			etMunschExtruder :=  ET_MunschExtruder_eError;             (* Next step *)
		END_IF

	ET_MunschExtruder_eSetCMD:
		tonWatchdog(
			IN := TRUE,
			PT:= tTimeOutAir
		);

		IF tonWatchdog.Q
		THEN
			tonWatchdog(IN := FALSE);

			bExtruderAirOn := FALSE;

			udnErrorNo := 1;

			etMunschExtruder := ET_MunschExtruder_eError;             (* Next step *)

		ELSIF bExtruderAirOn
		THEN
			IF bExtruderAirOk
			THEN
				tonWatchdog(IN := FALSE);

				etMunschExtruder := ET_MunschExtruder_eSetMaterialTemp;              (* Next step *)
			END_IF
		ELSE
			Munsch.stMunschCmd.etCommand := ET_MUNSCH_CMD_STOPHEAT;

			tonWatchdog(IN := FALSE);

			etMunschExtruder := ET_MunschExtruder_eExecuteCMD;              (* Next step *)
		END_IF

	ET_MunschExtruder_eSetMaterialTemp:
		nWatchdog := nWatchdog + 1;

		Munsch.bLockedInterface := FALSE;

		fbMaterialTemp(
			bEnable := TRUE,
			bExecute := TRUE,
			nMaterialTemp := nMaterialTemp,
			nMinMaterialTemp := nMinMaterialTemp,
			nMaxMaterialTemp := nMaxMaterialTemp,
			Munsch := Munsch
		);

		IF (NOT fbMaterialTemp.bBusy
		     AND fbMaterialTemp.bError)
		     OR nWatchdog > 1000
		THEN
			fbMaterialTemp(
				bEnable := TRUE,
				bExecute := FALSE,
				Munsch := Munsch
			);

			udnErrorNo := 2;                     (* Error number *)

			etMunschExtruder := ET_MunschExtruder_eError;             (* Next step *)
		
		ELSIF NOT fbMaterialTemp.bBusy
			   AND  fbMaterialTemp.bDone
		THEN
			fbMaterialTemp(
				bEnable := TRUE,
				bExecute := FALSE,
				Munsch := Munsch
			);

			nWatchdog := 0;

			etMunschExtruder := ET_MunschExtruder_eSetAirTemp;             (* Next step *)

		END_IF;

		Munsch.bLockedInterface := TRUE;
		Munsch.bReadStatus := FALSE;

	ET_MunschExtruder_eSetAirTemp:
		nWatchdog := nWatchdog + 1;

		Munsch.bLockedInterface := FALSE;

		fbAirTemp(
			bEnable := TRUE,
			bExecute := TRUE,
			nAirTemp := nAirTemp,
			nMinAirTemp := nMinAirTemp,
			nMaxAirTemp := nMaxAirTemp,
			Munsch := Munsch
		);

		IF (NOT fbAirTemp.bBusy
		     AND fbAirTemp.bError)
		     OR nWatchdog > 1000
		THEN
			fbAirTemp(
				bEnable := TRUE,
				bExecute := FALSE,
				Munsch := Munsch
			);

			udnErrorNo := 3;                     (* Error number *)

			etMunschExtruder := ET_MunschExtruder_eError;             (* Next step *)

		ELSIF NOT fbAirTemp.bBusy
			   AND fbAirTemp.bDone
		THEN
			fbAirTemp(
				bEnable := TRUE,
				bExecute := FALSE,
				Munsch := Munsch
			);

			nWatchdog := 0;

			Munsch.stMunschCmd.etCommand := ET_MUNSCH_CMD_STARTHEAT;

			etMunschExtruder := ET_MunschExtruder_eExecuteCMD;             (* Next step *)
		
		END_IF;

		Munsch.bLockedInterface := TRUE;
		Munsch.bReadStatus := FALSE;

	ET_MunschExtruder_eExecuteCMD:
		nWatchdog := nWatchdog + 1;

		Munsch.bSendExe := TRUE;

		IF Munsch.bStringReceived
		THEN
			IF (bExtruderAirOn
			      AND Munsch.stMunschRes.etResponse = ET_MUNSCH_RES_STARTHEAT)
			     OR
			     (NOT bExtruderAirOn
			      AND Munsch.stMunschRes.etResponse = ET_MUNSCH_RES_STOPHEAT)
			THEN
				Munsch.bSendExe := FALSE;

				nWatchdog := 0;

				etMunschExtruder := ET_MunschExtruder_eSetREQ;              (* Next step *)

			END_IF

		ELSIF Munsch.bInterfaceError
			    OR nWatchdog > 1000
		THEN
			Munsch.bSendExe := FALSE;

			udnErrorNo := 4;                     (* Error number *)

			etMunschExtruder := ET_MunschExtruder_eError;              (* Next step *)

		END_IF

	ET_MunschExtruder_eSetREQ:
		Munsch.stMunschCmd.etCommand := ET_MUNSCH_CMD_REQHEATSTATUS;

		etMunschExtruder := ET_MunschExtruder_eExecuteREQ;              (* Next step *)

	ET_MunschExtruder_eExecuteREQ:
		nWatchdog := nWatchdog + 1;

		Munsch.bSendExe := TRUE;

		IF Munsch.bStringReceived
		THEN
			IF Munsch.stMunschRes.etResponse = ET_MUNSCH_RES_ACKHEATSTATUSON
			THEN
				Munsch.bHeat := TRUE;
				Munsch.bSendExe := FALSE;

				nWatchdog := 0;
				etMunschExtruder := ET_MunschExtruder_eDone;              (* Next step *)
			
			ELSIF Munsch.stMunschRes.etResponse = ET_MUNSCH_RES_ACKHEATSTATUSOFF
			THEN
				Munsch.bHeat := FALSE;
				Munsch.bSendExe := FALSE;

				nWatchdog := 0;
				etMunschExtruder := ET_MunschExtruder_eDone;              (* Next step *)

			END_IF

		ELSIF Munsch.bInterfaceError
			    OR nWatchdog > 1000
		THEN
			Munsch.bSendExe := FALSE;

			udnErrorNo := 5;                     (* Error number *)

			etMunschExtruder := ET_MunschExtruder_eError;              (* Next step *)

		END_IF

	ET_MunschExtruder_eError:
		bBusy := FALSE;						(* Command busy *)
		bError := TRUE;						(* Command error  *)

		etMunschExtruder := ET_MunschExtruder_eNoExecute;

	ET_MunschExtruder_eDone:
		bDone := TRUE;						(* Command done *)
		bBusy := FALSE;						(* Command busy *)

		etMunschExtruder := ET_MunschExtruder_eNoExecute;

	ET_MunschExtruder_eNoExecute:
		IF NOT bStart
		     AND NOT bStop
		THEN
			(* Reset outputs *)
			bDone := FALSE;						(* Command done *)
			bBusy := FALSE;						(* Command busy *)
			bError := FALSE;						(* Command error  *)

			nWatchdog := 0;
			Munsch.bLockedInterface := FALSE;

			Munsch.stMunschCmd.etCommand := ET_MUNSCH_CMD_NOCMD;
			Munsch.stMunschRes.etResponse := ET_MUNSCH_RES_NOCMD;

			etMunschExtruder := ET_MunschExtruder_eWaitExecute;
		END_IF
END_CASE;

END_FUNCTION_BLOCK

// ---- POUs/Tc3 Objects/ExternalHardware/Munsch/FB_MunschExtruder_MaterialTemp_1.TcPOU
FUNCTION_BLOCK FB_MunschExtruder_MaterialTemp_1
(*

The function block used to control set material temperature on munschs extruder

Constructor: 		Patryk Panylo
Company:		E. Riexinger GmbH
Date:			18.10.2015
Version:			1.00

Date:			Revision:		Who:				Comment
dd.mm.yyyy		x.xx			Initials			comment

*)
VAR_INPUT
	(* Input variables / Eingang Variablen *)
	bEnable						:BOOL;						(* Enable FB signal *)
	bExecute					:BOOL;						(* Execut the function block *)
	nMaterialTemp				:INT;						(* Material temperatur *)
	nMinMaterialTemp			:INT;						(* Minimal material temperatur *)
	nMaxMaterialTemp			:INT;						(* Maximal material temperatur *)
	nMaterialTempTolerance		:INT := 5;						(* Material temperatur tolerance*)
END_VAR
VAR_OUTPUT
	(* Output variables / Ausgang Variablen *)
	bMaterialTempAlarm			:BOOL;						(* Exceeded material temperature tolerance  *)
	bDone						:BOOL;						(* Program done *)
	bBusy						:BOOL;						(* Program busy *)
	bError						:BOOL;						(* Error *)
	udnErrorNo					:UDINT;
END_VAR
VAR_IN_OUT
	(* Input Output variables / Ausgang Variablen *)
	Munsch						:ST_MUNSCH_REF;
END_VAR
VAR
	(* Enummerations *)
	etMunschExtruder				:ET_MunschExtruder;

	(* Variables *)
	nWatchdog					:INT;

	(* References *)

	(* Interfaces *)

	(* Instances *)
	rtExecute						:R_TRIG;

END_VAR

IF NOT bEnable
THEN
	bDone := FALSE;					(* Program done *)
	bBusy := FALSE;                                  	(* Program not busy *)
	bError := FALSE;                                 	(* Program not error *)
	udnErrorNo := 0;                                 		(* Error number *)

	RETURN;
END_IF;

(* Wait for triger *)
rtExecute(CLK := bExecute);

(* Send command *)
CASE etMunschExtruder OF

	ET_MunschExtruder_eWaitExecute:
		IF rtExecute.Q
		THEN
			nWatchdog := 0;

			Munsch.bSetAirTemp := FALSE;
			Munsch.bSetMaterialTemp := TRUE;
			Munsch.bStartHeat := FALSE;
			Munsch.bStopHeat  := FALSE;
			Munsch.bStartExtruding := FALSE;
			Munsch.bStopExtruding  := FALSE;
			Munsch.bReadStatus := FALSE;

			etMunschExtruder := ET_MunschExtruder_eChkInterface;              (* Next step *)
		END_IF

	ET_MunschExtruder_eChkInterface:
		nWatchdog := nWatchdog + 1;

		IF NOT Munsch.bLockedInterface
		THEN
			bBusy := FALSE;                                     	(* Program not busy *)
			bError := FALSE;                         		(* Program not error *)
			udnErrorNo := 0;                         		(* Error number *)

			IF Munsch.bSetMaterialTemp
			THEN
				nWatchdog := 0;
				bDone:= FALSE;                               		(* Program done *)
				bBusy := TRUE;                                  	(* Program busy *)
	
				Munsch.bLockedInterface := TRUE;
				Munsch.bSendExe := FALSE;
	
				IF nMaterialTemp >= nMinMaterialTemp
				     AND nMaterialTemp <= nMaxMaterialTemp
				THEN
					etMunschExtruder := ET_MunschExtruder_eSetCMD;              (* Next step *)
				ELSE
					udnErrorNo := 1;
	
					etMunschExtruder := ET_MunschExtruder_eError;              (* Next step *)
				END_IF

			ELSE
				etMunschExtruder := ET_MunschExtruder_eError;             (* Next step *)
			END_IF

			Munsch.bSetMaterialTemp := FALSE;

		ELSIF nWatchdog > 1000
		THEN
			Munsch.bSetMaterialTemp := FALSE;

			etMunschExtruder := ET_MunschExtruder_eError;             (* Next step *)
		END_IF

	ET_MunschExtruder_eSetCMD:
		Munsch.stMunschCmd.etCommand := ET_MUNSCH_CMD_SETMATERIALTEMP;
		Munsch.stMunschCmd.nMaterialTemp := nMaterialTemp;

		etMunschExtruder := ET_MunschExtruder_eExecuteCMD;              (* Next step *)

	ET_MunschExtruder_eExecuteCMD:
		nWatchdog := nWatchdog + 1;

		Munsch.bSendExe := TRUE;

		IF Munsch.bStringReceived
		THEN
			IF Munsch.stMunschRes.etResponse = ET_MUNSCH_RES_SETMATERIALTEMP
			     AND Munsch.stMunschCmd.nMaterialTemp = Munsch.stMunschRes.nMaterialRefTemp
			THEN
				Munsch.bSendExe := FALSE;

				nWatchdog := 0;
				etMunschExtruder := ET_MunschExtruder_eSetREQ;              (* Next step *)
			END_IF

		ELSIF Munsch.bInterfaceError
			    OR nWatchdog > 1000
		THEN
			Munsch.bSendExe := FALSE;

			udnErrorNo := 2;                     (* Error number *)
			etMunschExtruder := ET_MunschExtruder_eError;              (* Next step *)
		END_IF

	ET_MunschExtruder_eSetREQ:
		Munsch.stMunschCmd.etCommand := ET_MUNSCH_CMD_REQMATERIALREFTEMP;

		etMunschExtruder := ET_MunschExtruder_eExecuteREQ;              (* Next step *)

	ET_MunschExtruder_eExecuteREQ:
		nWatchdog := nWatchdog + 1;

		Munsch.bSendExe := TRUE;

		IF Munsch.bStringReceived
		THEN
			IF Munsch.stMunschRes.etResponse = ET_MUNSCH_RES_REQMATERIALREFTEMP
			THEN
				Munsch.nMaterialRefTemp := Munsch.stMunschRes.nMaterialRefTemp;

				Munsch.bSendExe := FALSE;

				nWatchdog := 0;
				etMunschExtruder := ET_MunschExtruder_eDone;              (* Next step *)

			END_IF

		ELSIF Munsch.bInterfaceError
			    OR nWatchdog > 1000
		THEN
			Munsch.bSendExe := FALSE;

			udnErrorNo := 3;                     (* Error number *)
			etMunschExtruder := ET_MunschExtruder_eError;              (* Next step *)
		END_IF

	ET_MunschExtruder_eError:
		bBusy := FALSE;						(* Command busy *)
		bError := TRUE;						(* Command error  *)

		etMunschExtruder := ET_MunschExtruder_eNoExecute;

	ET_MunschExtruder_eDone:
		bDone := TRUE;						(* Command done *)
		bBusy := FALSE;						(* Command busy *)

		etMunschExtruder := ET_MunschExtruder_eNoExecute;

	ET_MunschExtruder_eNoExecute:
		IF NOT bExecute
		THEN
			(* Reset outputs *)
			bDone := FALSE;						(* Command done *)
			bBusy := FALSE;						(* Command busy *)
			bError := FALSE;						(* Command error  *)

			nWatchdog := 0;
			Munsch.bLockedInterface := FALSE;

			Munsch.stMunschCmd.etCommand := ET_MUNSCH_CMD_NOCMD;
			Munsch.stMunschRes.etResponse := ET_MUNSCH_RES_NOCMD;

			etMunschExtruder := ET_MunschExtruder_eWaitExecute;
		END_IF
END_CASE;

bMaterialTempAlarm := Munsch.nMaterialActTemp > Munsch.nMaterialRefTemp + nMaterialTempTolerance
					 OR Munsch.nMaterialActTemp > Munsch.nMaterialRefTemp - nMaterialTempTolerance;

END_FUNCTION_BLOCK

// ---- POUs/Tc3 Objects/ExternalHardware/Munsch/FB_MunschExtruder_ReadStatus_1.TcPOU
FUNCTION_BLOCK FB_MunschExtruder_ReadStatus_1
(*

The function block used to read status of Munsch extruder

Constructor: 		Patryk Panylo
Company:		E. Riexinger GmbH
Date:			13.10.2015
Version:			1.00

Date:			Revision:		Who:				Comment
dd.mm.yyyy		x.xx			Initials			comment

*)
VAR_INPUT
	(* Input variables / Eingang Variablen *)
	bEnable						:BOOL;						(* Enable FB signal *)
	bExecute					:BOOL;						(* Execute read status *)
	tReadStatus					:TIME := t#0ms;				(* Read current status *)
END_VAR
VAR_OUTPUT
	(* Output variables / Ausgang Variablen *)
	bDone						:BOOL;						(* Program done *)
	bBusy						:BOOL;						(* Program busy *)
	bError						:BOOL;						(* Error *)
	udnErrorNo					:UDINT;
END_VAR
VAR_IN_OUT
	(* Input Output variables / Ausgang Variablen *)
	Munsch						:ST_MUNSCH_REF;
END_VAR
VAR
	(* Enummerations *)
	etMunschExtruder				:ET_MunschExtruder;

	(* Variables *)
	bReadStatus					:BOOL;
	nReqCount					:INT;
	nWatchdog					:INT;

	(* References *)

	(* Interfaces *)

	(* Instances *)
	tonReadStatus				:TON;
	rtExecute						:R_TRIG;
	rtStart						:R_TRIG;
	rtStop						:R_TRIG;
END_VAR

IF NOT bEnable
THEN
	bDone := FALSE;					(* Program done *)
	bBusy := FALSE;                                  	(* Program not busy *)
	bError := FALSE;                                 	(* Program not error *)
	udnErrorNo := 0;                                 		(* Error number *)

	tonReadStatus(
		IN := FALSE,
	);

	RETURN;
END_IF;

rtStart(CLK := (tReadStatus > t#0ms
		       OR  (bExecute AND tReadStatus = t#0ms))
		       AND NOT Munsch.bLockedInterface);
rtStop(CLK := tReadStatus = t#0ms);

IF rtStop.Q
THEN
	Munsch.bReadStatus := FALSE;

ELSIF rtStart.Q
THEN
	Munsch.bReadStatus := TRUE;

	bDone := FALSE;					(* Program done *)
	bBusy := FALSE;                                  	(* Program not busy *)
	bError := FALSE;                                 	(* Program not error *)
	udnErrorNo := 0;                                 		(* Error number *)

	etMunschExtruder := ET_MunschExtruder_eWaitExecute;              (* Next step *)

END_IF

tonReadStatus(
	IN := Munsch.bReadStatus,
	PT := tReadStatus,
);

rtExecute(
	CLK := tonReadStatus.Q
);

(* Send command *)
CASE etMunschExtruder OF

	ET_MunschExtruder_eWaitExecute:
		bBusy := FALSE;                                     	(* Program not busy *)
		bError := FALSE;                         		(* Program not error *)
		udnErrorNo := 0;                         		(* Error number *)

		IF rtExecute.Q
		     AND NOT Munsch.bLockedInterface
		THEN
			nWatchdog := 0;
			bDone:= FALSE;                               		(* Program done *)
			bBusy := TRUE;                                  	(* Program busy *)

			nReqCount  := 0;
			Munsch.bLockedInterface := TRUE;
			Munsch.bSendExe := FALSE;

			etMunschExtruder := ET_MunschExtruder_eSetREQ;              (* Next step *)

		END_IF

	ET_MunschExtruder_eSetREQ:
		CASE nReqCount
		OF
			0: Munsch.stMunschCmd.etCommand := ET_MUNSCH_CMD_REQHEATSTATUS;
			    nReqCount := 1;
			1: Munsch.stMunschCmd.etCommand := ET_MUNSCH_CMD_REQEXTRUDERSTATUS;
			    nReqCount := 2;
			2: Munsch.stMunschCmd.etCommand := ET_MUNSCH_CMD_REQMATERIALREFTEMP;
			    nReqCount := 3;
			3: Munsch.stMunschCmd.etCommand := ET_MUNSCH_CMD_REQMATERIALACTTEMP;
			    nReqCount := 4;
			4: Munsch.stMunschCmd.etCommand := ET_MUNSCH_CMD_REQAIRREFTEMP;
			    nReqCount := 5;
			5: Munsch.stMunschCmd.etCommand := ET_MUNSCH_CMD_REQAIRACTTEMP;
			    nReqCount := 6;
			6: Munsch.stMunschCmd.etCommand := ET_MUNSCH_CMD_REQSTATUS;
				nReqCount := 0;
		END_CASE

		etMunschExtruder := ET_MunschExtruder_eExecuteREQ;              (* Next step *)

	ET_MunschExtruder_eExecuteREQ:
		nWatchdog := nWatchdog + 1;

		Munsch.bSendExe := TRUE;

		IF Munsch.bStringReceived
		THEN
			IF Munsch.stMunschRes.etResponse = ET_MUNSCH_RES_ACKHEATSTATUSON
			THEN
				Munsch.bHeat := TRUE;
				Munsch.bSendExe := FALSE;

				nWatchdog := 0;
				IF nReqCount > 0
				     AND Munsch.bReadStatus
				THEN
					etMunschExtruder := ET_MunschExtruder_eSetREQ;
				ELSE
					etMunschExtruder := ET_MunschExtruder_eDone;              (* Next step *)
				END_IF
			
			ELSIF Munsch.stMunschRes.etResponse = ET_MUNSCH_RES_ACKHEATSTATUSOFF
			THEN
				Munsch.bHeat := FALSE;
				Munsch.bSendExe := FALSE;

				nWatchdog := 0;
				IF nReqCount > 0
				    AND Munsch.bReadStatus
				THEN
					etMunschExtruder := ET_MunschExtruder_eSetREQ;
				ELSE
					etMunschExtruder := ET_MunschExtruder_eDone;              (* Next step *)
				END_IF

			ELSIF Munsch.stMunschRes.etResponse = ET_MUNSCH_RES_ACKEXTRUDERSTATUSON
			THEN
				Munsch.bExtruding := TRUE;
				Munsch.bSendExe := FALSE;

				nWatchdog := 0;
				IF nReqCount > 0
				    AND Munsch.bReadStatus
				THEN
					etMunschExtruder := ET_MunschExtruder_eSetREQ;
				ELSE
					etMunschExtruder := ET_MunschExtruder_eDone;              (* Next step *)
				END_IF
			
			ELSIF Munsch.stMunschRes.etResponse = ET_MUNSCH_RES_ACKEXTRUDERSTATUSOFF
			THEN
				Munsch.bExtruding := FALSE;
				Munsch.bSendExe := FALSE;

				nWatchdog := 0;
				IF nReqCount > 0
				     AND Munsch.bReadStatus
				THEN
					etMunschExtruder := ET_MunschExtruder_eSetREQ;
				ELSE
					etMunschExtruder := ET_MunschExtruder_eDone;              (* Next step *)
				END_IF

			ELSIF Munsch.stMunschRes.etResponse = ET_MUNSCH_RES_REQMATERIALREFTEMP
			THEN
				Munsch.nMaterialRefTemp := Munsch.stMunschRes.nMaterialRefTemp;
				Munsch.bSendExe := FALSE;

				nWatchdog := 0;
				IF nReqCount > 0
				     AND Munsch.bReadStatus
				THEN
					etMunschExtruder := ET_MunschExtruder_eSetREQ;
				ELSE
					etMunschExtruder := ET_MunschExtruder_eDone;              (* Next step *)
				END_IF

			ELSIF Munsch.stMunschRes.etResponse = ET_MUNSCH_RES_REQMATERIALACTTEMP
			THEN
				Munsch.nMaterialActTemp := Munsch.stMunschRes.nMaterialActTemp;
				Munsch.bSendExe := FALSE;

				nWatchdog := 0;
				IF nReqCount > 0
				     AND Munsch.bReadStatus
				THEN
					etMunschExtruder := ET_MunschExtruder_eSetREQ;
				ELSE
					etMunschExtruder := ET_MunschExtruder_eDone;              (* Next step *)
				END_IF

			ELSIF Munsch.stMunschRes.etResponse = ET_MUNSCH_RES_REQAIRREFTEMP
			THEN
				Munsch.nAirRefTemp := Munsch.stMunschRes.nAirRefTemp;
				Munsch.bSendExe := FALSE;

				nWatchdog := 0;
				IF nReqCount > 0
				     AND Munsch.bReadStatus
				THEN
					etMunschExtruder := ET_MunschExtruder_eSetREQ;
				ELSE
					etMunschExtruder := ET_MunschExtruder_eDone;              (* Next step *)
				END_IF

			ELSIF Munsch.stMunschRes.etResponse = ET_MUNSCH_RES_REQAIRACTTEMP
			THEN
				Munsch.nAirActTemp := Munsch.stMunschRes.nAirActTemp;
				Munsch.bSendExe := FALSE;

				nWatchdog := 0;
				IF nReqCount > 0
				     AND Munsch.bReadStatus
				THEN
					etMunschExtruder := ET_MunschExtruder_eSetREQ;
				ELSE
					etMunschExtruder := ET_MunschExtruder_eDone;              (* Next step *)
				END_IF

			ELSIF Munsch.stMunschRes.etResponse = ET_MUNSCH_RES_REQSTATUSHEATED
			THEN
				Munsch.bHeating := FALSE;
				Munsch.bHeated := TRUE;
				Munsch.bError := FALSE;
				Munsch.bSendExe := FALSE;

				nWatchdog := 0;
				IF nReqCount > 0
				     AND Munsch.bReadStatus
				THEN
					etMunschExtruder := ET_MunschExtruder_eSetREQ;
				ELSE
					etMunschExtruder := ET_MunschExtruder_eDone;              (* Next step *)
				END_IF

			ELSIF Munsch.stMunschRes.etResponse = ET_MUNSCH_RES_REQSTATUSHEATING
			THEN
				Munsch.bHeating := Munsch.bHeat;
				Munsch.bHeated := FALSE;
				Munsch.bError := FALSE;
				Munsch.bSendExe := FALSE;

				nWatchdog := 0;
				IF nReqCount > 0
				     AND Munsch.bReadStatus
				THEN
					etMunschExtruder := ET_MunschExtruder_eSetREQ;
				ELSE
					etMunschExtruder := ET_MunschExtruder_eDone;              (* Next step *)
				END_IF

			ELSIF Munsch.stMunschRes.etResponse = ET_MUNSCH_RES_REQSTATUSERROR
			THEN
				Munsch.bHeating := FALSE;
				Munsch.bHeated := FALSE;
				Munsch.bError := TRUE;
				Munsch.bSendExe := FALSE;

				nWatchdog := 0;
				IF nReqCount > 0
				     AND Munsch.bReadStatus
				THEN
					etMunschExtruder := ET_MunschExtruder_eSetREQ;
				ELSE
					etMunschExtruder := ET_MunschExtruder_eDone;              (* Next step *)
				END_IF

			END_IF

		ELSIF Munsch.bInterfaceError
 			    OR nWatchdog > 1000
		THEN
			Munsch.bSendExe := FALSE;

			udnErrorNo := 2;                     (* Error number *)

			etMunschExtruder := ET_MunschExtruder_eError;              (* Next step *)
		END_IF

	ET_MunschExtruder_eError:
		bBusy := FALSE;						(* Command busy *)
		bError := TRUE;						(* Command error  *)

		etMunschExtruder := ET_MunschExtruder_eNoExecute;

	ET_MunschExtruder_eDone:
		bDone := TRUE;						(* Command done *)
		bBusy := FALSE;						(* Command busy *)

		etMunschExtruder := ET_MunschExtruder_eNoExecute;

	ET_MunschExtruder_eNoExecute:
		IF tReadStatus > t#0ms
		THEN
			tonReadStatus(
				IN := FALSE,
				PT := tReadStatus,
			);
		END_IF

		IF NOT tonReadStatus.Q
		     OR (NOT bExecute AND tReadStatus = t#0ms)
		THEN
			(* Reset outputs *)
			bDone := FALSE;						(* Command done *)
			bBusy := FALSE;						(* Command busy *)
			bError := FALSE;						(* Command error  *)

			nWatchdog := 0;
			Munsch.bLockedInterface := FALSE;

			IF tReadStatus = t#0ms
			THEN
				Munsch.bReadStatus := FALSE;
			END_IF

			etMunschExtruder := ET_MunschExtruder_eWaitExecute;
		END_IF
END_CASE;

END_FUNCTION_BLOCK

// ---- POUs/Tc3 Objects/ExternalHardware/Munsch/FB_MUNSCH_EXTRUDER_REF_1.TcPOU
FUNCTION_BLOCK FB_MUNSCH_EXTRUDER_REF_1
VAR_INPUT
	bSendExe					:BOOL;						(* Send execute *)
	tSendPeriod					:TIME := t#0s;					(* Send data every period. If tSendPeriod is 0 then th function is not active *)
	bLockedInterface				:BOOL;						(* Locked interface *)
	bHeat						:BOOL;						(* Heat status ON = TRUE, OFF = FALSE *)
	bHeating						:BOOL;						(* Heating status ON = TRUE, OFF = FALSE *)
	bHeated						:BOOL;						(* Heated status ON = TRUE, OFF = FALSE *)
	bError						:BOOL;						(* Error ON = TRUE, OFF = FALSE *)
	bExtruding					:BOOL;						(* Extruder status ON = TRUE, OFF = FALSE *)
	nMaterialRefTemp			:INT;						(* Referenc material tamperature *)
	nMaterialActTemp				:INT;						(* Current material tamperature *)
	nAirRefTemp					:INT;						(* Referenc air tamperature *)
	nAirActTemp					:INT;						(* Current air tamperature *)
	stMunschCmd				:ST_MUNSCH_CMD_Data;
	stMunschRes					:ST_MUNSCH_RES_Data;
	bInterfaceReady				:BOOL;						(* Interface ready to use *)
	bInterfaceError				:BOOL;						(* Interface error *)
	bStringReceived				:BOOL;						(* String received *)
	bSetAirTemp					:BOOL;						(* Set air temperature *)
	bSetMaterialTemp			:BOOL;						(* Set material temperature *)
	bStartHeat					:BOOL;						(* Heat start *)
	bStopHeat					:BOOL;						(* Heat stop *)
	bStartExtruding				:BOOL;						(* Extruding start *)
	bStopExtruding				:BOOL;						(* Extruding start *)
	bReadStatus					:BOOL;						(* Enable read current status *)
	bExtrudingStop				:BOOL;						(* Extruding stop *)
	nExtrudingSpeed				:INT;						(* Extruding speed *)
END_VAR
VAR_OUTPUT

END_VAR
VAR_IN_OUT

END_VAR
VAR

END_VAR

;

END_FUNCTION_BLOCK

// ---- POUs/Tc3 Objects/ExternalHardware/Munsch/F_MunschCMD_1.TcPOU
FUNCTION F_MunschCMD_1 : STRING							(* Command to Munsch extruder *)
VAR_INPUT
	stMunschCmd			:ST_MUNSCH_CMD_Data;
END_VAR
VAR
	usnBaseMaterialTemp		:USINT := 160;					(* Base material temperature 160 °C *)
	usnBaseAirTemp			:USINT := 160;					(* Base air temperature 160 °C *)
END_VAR


CASE stMunschCmd.etCommand OF

	ET_MUNSCH_CMD_NOCMD:						F_MunschCMD := 'NoCmd';
	ET_MUNSCH_CMD_STARTHEAT:					F_MunschCMD := 'H1';
	ET_MUNSCH_CMD_STOPHEAT:					F_MunschCMD := 'H0';
	ET_MUNSCH_CMD_REQHEATSTATUS:			F_MunschCMD := 'h?';
	ET_MUNSCH_CMD_STARTEXTRUDER:			F_MunschCMD := 'R1';
	ET_MUNSCH_CMD_STOPEXTRUDER:				F_MunschCMD := 'R0';
	ET_MUNSCH_CMD_REQEXTRUDERSTATUS:		F_MunschCMD := 'r?';
	ET_MUNSCH_CMD_SETMATERIALTEMP:			F_MunschCMD := CONCAT('M', CHR(INT_TO_BYTE(MIN(MAX(stMunschCmd.nMaterialTemp - usnBaseMaterialTemp, 0), 240))));
	ET_MUNSCH_CMD_REQMATERIALREFTEMP:		F_MunschCMD := 'm?';
	ET_MUNSCH_CMD_REQMATERIALACTTEMP:		F_MunschCMD := 'n?';
	ET_MUNSCH_CMD_SETAIRTEMP:					F_MunschCMD := CONCAT('A', CHR(INT_TO_BYTE(MIN(MAX(stMunschCmd.nAirTemp - usnBaseAirTemp, 0), 240))));
	ET_MUNSCH_CMD_REQAIRREFTEMP:				F_MunschCMD := 'a?';
	ET_MUNSCH_CMD_REQAIRACTTEMP:				F_MunschCMD := 'b?';
	ET_MUNSCH_CMD_REQSTATUS:					F_MunschCMD := 's?';
ELSE
	F_MunschCMD := 'NoCmd';
END_CASE

END_FUNCTION

// ---- POUs/Tc3 Objects/ExternalHardware/Munsch/F_MunschRES_1.TcPOU
FUNCTION F_MunschRES_1 : ST_MUNSCH_RES_Data			(* Response from Munsch extruder *)
VAR_INPUT
	sResponse					:STRING	;
END_VAR
VAR
	usnBaseMaterialTemp		:USINT := 160;					(* Base material temperature 160 °C *)
	usnBaseAirTemp			:USINT := 160;					(* Base air temperature 160 °C *)
END_VAR


IF sResponse = 'H1'		THEN	F_MunschRES.etResponse := ET_MUNSCH_RES_STARTHEAT;
ELSIF sResponse = 'H0'	THEN	F_MunschRES.etResponse := ET_MUNSCH_RES_STOPHEAT;
ELSIF sResponse = 'h1'	THEN	F_MunschRES.etResponse := ET_MUNSCH_RES_ACKHEATSTATUSON;
ELSIF sResponse = 'h0'	THEN	F_MunschRES.etResponse := ET_MUNSCH_RES_ACKHEATSTATUSOFF;
ELSIF sResponse = 'R1'	THEN	F_MunschRES.etResponse := ET_MUNSCH_RES_STARTEXTRUDER;
ELSIF sResponse = 'R0'	THEN	F_MunschRES.etResponse := ET_MUNSCH_RES_STOPEXTRUDER;
ELSIF sResponse = 'r1'		THEN	F_MunschRES.etResponse := ET_MUNSCH_RES_ACKEXTRUDERSTATUSON;
ELSIF sResponse = 'r0'		THEN	F_MunschRES.etResponse := ET_MUNSCH_RES_ACKEXTRUDERSTATUSOFF;
ELSIF FIND(sResponse, 'M') = 1		THEN	F_MunschRES.etResponse := ET_MUNSCH_RES_SETMATERIALTEMP; F_MunschRES.nMaterialRefTemp := usnBaseMaterialTemp + ASC(DELETE(sResponse,LEN('M'), FIND(sResponse, 'M')));
ELSIF FIND(sResponse, 'm') = 1 		THEN	F_MunschRES.etResponse := ET_MUNSCH_RES_REQMATERIALREFTEMP; F_MunschRES.nMaterialRefTemp := usnBaseMaterialTemp + ASC(DELETE(sResponse,LEN('m'), FIND(sResponse, 'm')));
ELSIF FIND(sResponse, 'n') = 1 		THEN	F_MunschRES.etResponse := ET_MUNSCH_RES_REQMATERIALACTTEMP; F_MunschRES.nMaterialActTemp := usnBaseMaterialTemp + ASC(DELETE(sResponse,LEN('n'), FIND(sResponse, 'n')));
ELSIF FIND(sResponse, 'A') = 1		THEN	F_MunschRES.etResponse := ET_MUNSCH_RES_SETAIRTEMP; F_MunschRES.nAirRefTemp := usnBaseAirTemp + ASC(DELETE(sResponse,LEN('A'), FIND(sResponse, 'A')));
ELSIF FIND(sResponse, 'a') = 1		THEN	F_MunschRES.etResponse := ET_MUNSCH_RES_REQAIRREFTEMP; F_MunschRES.nAirRefTemp := usnBaseAirTemp + ASC(DELETE(sResponse,LEN('a'), FIND(sResponse, 'a')));
ELSIF FIND(sResponse, 'b') = 1		THEN	F_MunschRES.etResponse := ET_MUNSCH_RES_REQAIRACTTEMP; F_MunschRES.nAirActTemp := usnBaseAirTemp + ASC(DELETE(sResponse,LEN('b'), FIND(sResponse, 'b')));
ELSIF sResponse = 's1'	THEN	F_MunschRES.etResponse := ET_MUNSCH_RES_REQSTATUSHEATED;
ELSIF sResponse = 's0'	THEN	F_MunschRES.etResponse := ET_MUNSCH_RES_REQSTATUSHEATING;
ELSIF sResponse = 'sE'	THEN	F_MunschRES.etResponse := ET_MUNSCH_RES_REQSTATUSERROR;
ELSIF sResponse = 'ER' 	THEN	F_MunschRES.etResponse := ET_MUNSCH_RES_CMDERROR;
ELSE F_MunschRES.etResponse := ET_MUNSCH_RES_NOCMD;
END_IF

END_FUNCTION

// ---- POUs/Tc3 Objects/ExternalHardware/Periphery/FB_PERIPHERY_REF_1.TcPOU
FUNCTION_BLOCK FB_PERIPHERY_REF_1
VAR_INPUT

END_VAR
VAR_OUTPUT

END_VAR
VAR_IN_OUT

END_VAR
VAR

END_VAR

;

END_FUNCTION_BLOCK

// ---- POUs/Tc3 Objects/ExternalHardware/YASKAWA/FB_YASKAWA_Controller_1.TcPOU
FUNCTION_BLOCK FB_YASKAWA_Controller_1
(*

The function block used to control axis.

Constructor: 		Patryk Panylo
Company:		E. Riexinger GmbH
Date:			20.06.2018
Version:			1.00

Date:			Revision:		Who:				Comment
dd.mm.yyyy		x.xx			Initials			comment

*)
VAR_INPUT
	(* Input variables / Eingang Variablen *)
	bEnable						:BOOL;						(* Signal FB enable *)
	etMachineMode				:ET_MachineMode;			(* Machine mode *)
	etMachineState				:ET_MachineState;			(* Machine state *)
	bDrivesOn					:BOOL;						(* Enable the drives *)
	bMoveOn					:BOOL;						(* Enable the move enable *)
	bReset						:BOOL;						(* Signal reset *)
	bExeReset					:BOOL;						(* Execute auto reset *)
	lrOverride					:LREAL;						(* Override 100% percent *)
END_VAR
VAR_OUTPUT
	(* Output variables / Ausgang Variablen *)
	bStatus						:BOOL;						(* Feedback *)
	bStatusDelay					:BOOL;						(* Feedback delay *)
	bReseted					:BOOL;						(* Reset completed *)
	bError						:BOOL;						(* Controller error *)
	udnErrorNo					:UDINT;						(* Error number *)
	bInHome						:BOOL;						(* In home *)
	bNotMoving					:BOOL;						(* Status of moving *)
	bNotInCrashAreaMachine		:BOOL;						(* Status not in crash area *)
END_VAR
VAR_IN_OUT
	(* Input Output variables / Ausgang Variablen *)
	Yaskawa					:ST_YASKAWA_REF;				(* The YASKAWA_REF data type  is an interface between the PLC and the YASKAWA and contains axis information *)
END_VAR
VAR
	(* Enummerations *)

	(* Variables *)
	tStatusDelay					:TIME := t#1s;					(* Status delay time *)

	bFirstTime					:BOOL;

	(* References *)

	(* Interfaces *)

	(* Instances *)
	fbPower						:FB_YASKAWA_Power;		(* The function block is used to enable for an axis *)
	tonStatusDelay				:TON;						(* Delay controller enabled status *)
	fbReset						:FB_YASKAWA_Reset;			(* An axis reset is carried out with the function block *)

END_VAR


IF NOT bEnable							(* Signal FB enable *)
THEN
	bStatus := FALSE;						(* Feedback *)
	bStatusDelay := FALSE;				(* Feedback *)
	bError := FALSE;						(* Controller error *)
	udnErrorNo := 0;						(* Error number *)

	bFirstTime := FALSE;
	RETURN;
END_IF

IF NOT bFirstTime
THEN

	bFirstTime := TRUE;
END_IF;

A_Power();
A_Reset();
A_Error();

(* In home *)
bInHome := Yaskawa.stYaskawaToPlc.bInHome;

(* Status not moving *)
bNotMoving := Yaskawa.stYaskawaToPlc.bNotMoving;

(* Status not in crash area *)
bNotInCrashAreaMachine := Yaskawa.stYaskawaToPlc.bNotInCrashAreaMachine;

ACTION A_Error:

bError := fbReset.bError
	         OR fbPower.bError;
END_ACTION

ACTION A_Power:

fbPower(
	bEnable := TRUE,
	bAutoHand := etMachineMode = ET_MachineMode_eHome
			         OR etMachineMode = ET_MachineMode_eStepping
			         OR etMachineMode = ET_MachineMode_eAutomatic
					 OR etMachineMode = ET_MachineMode_eMaintenance,
	bDrivesOn :=  bDrivesOn,
	bMoveOn := bMoveOn,
	lrOverride := lrOverride,
	Yaskawa := Yaskawa
 );

tonStatusDelay(
	IN := fbPower.bStatus,
	PT := SEL(etMachineMode = ET_MachineMode_eManual, tStatusDelay, t#0ms),
	Q => bStatusDelay
);
END_ACTION

ACTION A_Reset:

fbReset(
	bExecute := bReset
	            	     XOR bExeReset,
	Yaskawa := Yaskawa,
	bDone => bReseted
);
END_ACTION

END_FUNCTION_BLOCK

// ---- POUs/Tc3 Objects/ExternalHardware/YASKAWA/FB_YASKAWA_Power_1.TcPOU
FUNCTION_BLOCK FB_YASKAWA_Power_1
(*

The function block used to enable drives for an yaskawa

Constructor: 		Patryk Panylo
Company:		E. Riexinger GmbH
Date:			20.06.2018
Version:			1.00

Date:			Revision:		Who:				Comment

*)
VAR_INPUT
	(* Input variables / Eingang Variablen *)
	bEnable						:BOOL;			(* Signal FB enable *)
	bAutoHand					:BOOL;			(* Auto := TRUE, Hand := FALSE *)
	bDrivesOn					:BOOL;			(* Enable the drives *)
	bMoveOn					:BOOL;			(* Enable the move enable *)
	lrOverride					:LREAL;			(* Velocity override in % for all motion commands. (0 <= Override <= 100.0) *)
END_VAR
VAR_OUTPUT
	(* Output variables / Ausgang Variablen *)
	bStatus						:BOOL;			(* Status = TRUE indicates that the axis is ready for operation. *)
	bError						:BOOL;			(* Error *)
	udnErrorNo					:UDINT;			(* Error number *)
	sErrorMsg					:STRING; 		(* Error message *)
END_VAR
VAR_IN_OUT
	(* Input Output variables / Ausgang Variablen *)
	Yaskawa					:ST_YASKAWA_REF;				(* The YASKAWA_REF data type  is an interface between the PLC and the YASKAWA and contains axis information *)
END_VAR
VAR
	(* Enummerations *)

	(* Variables *)
	tStatusDelay 					:TIME := t#300ms;

	(* References *)

	(* Interfaces *)

	(* Instances *)
	tonStatusDelay				:TON;
END_VAR


IF NOT bEnable
THEN
	Yaskawa.stPlcToYaskawa.bExternalServoOn := FALSE;                   		 (* Switch on *)
	tonStatusDelay(IN := FALSE,
				    PT := tStatusDelay);
ELSE

	IF NOT bDrivesOn
	     OR Yaskawa.stYaskawaToPlc.bAlarmErrorOccured
	THEN
		Yaskawa.stPlcToYaskawa.bCallMasterJob := FALSE;
		Yaskawa.stPlcToYaskawa.bExternalStart := FALSE;
		Yaskawa.stPlcToYaskawa.bExternalHold := FALSE;
		Yaskawa.stPlcToYaskawa.bExternalServoOn := FALSE;						 (* Switch on *)
		Yaskawa.stPlcToYaskawa.bExternalServoOffEStop := TRUE;                   		 (* Switch off *)
		Yaskawa.stPlcToYaskawa.bExternalServoOffHoldStop := FALSE;                   		 (* Switch off *)
	ELSE
		IF bAutoHand			(* Auto *)
		THEN
			IF bMoveOn
			     AND Yaskawa.stYaskawaToPlc.bRemoteModeSelected
			THEN
				Yaskawa.stPlcToYaskawa.bExternalServoOn := TRUE;                   				 (* Switch on *)
				Yaskawa.stPlcToYaskawa.bExternalServoOffEStop := FALSE;                   		 (* Switch off *)
				Yaskawa.stPlcToYaskawa.bExternalServoOffHoldStop := FALSE;                   		 (* Switch off *)
			ELSE
				Yaskawa.stPlcToYaskawa.bExternalServoOn := FALSE;                   				(* Switch on *)
				Yaskawa.stPlcToYaskawa.bExternalServoOffEStop := FALSE;                   		(* Switch off *)
				Yaskawa.stPlcToYaskawa.bExternalServoOffHoldStop := TRUE;				(* Switch off *)
			END_IF
		ELSE				(* Manual *)
			Yaskawa.stPlcToYaskawa.bCallMasterJob := FALSE;
			Yaskawa.stPlcToYaskawa.bExternalStart := FALSE;
			Yaskawa.stPlcToYaskawa.bExternalHold := FALSE;
			Yaskawa.stPlcToYaskawa.bExternalServoOn := FALSE;						(* Switch on *)
			Yaskawa.stPlcToYaskawa.bExternalServoOffEStop := FALSE;                   		(* Switch off *)
			Yaskawa.stPlcToYaskawa.bExternalServoOffHoldStop := FALSE;				(* Switch off *)
		END_IF
	END_IF;
END_IF;

Yaskawa.stPlcToYaskawa.nOverride := LREAL_TO_INT(LIMIT(0,lrOverride,100));

tonStatusDelay(IN := Yaskawa.stYaskawaToPlc.bServoIsOn,		(* Control enabled *)
			   PT := tStatusDelay);
bStatus := tonStatusDelay.Q;

END_FUNCTION_BLOCK

// ---- POUs/Tc3 Objects/ExternalHardware/YASKAWA/FB_YASKAWA_REF_1.TcPOU
FUNCTION_BLOCK FB_YASKAWA_REF_1
VAR_INPUT
	stYaskawaToPlc				:ST_YASKAWATOPLC;
	stPlcToYaskawa				:ST_PLCTOYASKAWA;

	stRobotToPlc					AT %I*:ST_ROBOTTOPLC;
	stPlcToRobot					AT %Q*:ST_PLCTOROBOT;
END_VAR
VAR_OUTPUT

END_VAR
VAR_IN_OUT

END_VAR
VAR

END_VAR

;

END_FUNCTION_BLOCK

// ---- POUs/Tc3 Objects/ExternalHardware/YASKAWA/FB_YASKAWA_Reset_1.TcPOU
FUNCTION_BLOCK FB_YASKAWA_Reset_1
(*

The function block used to reset the yaskawa message.

Constructor: 		Patryk Panylo
Company:		E. Riexinger GmbH
Date:			20.06.2018
Version:			1.00

Date:			Revision:		Who:				Comment

*)
VAR_INPUT
	(* Input variables / Eingang Variablen *)
	bExecute					:BOOL;		(* Execut the function block *)
	bExtReset					:BOOL;
END_VAR
VAR_OUTPUT
	(* Output variables / Ausgang Variablen *)
	bDone						:BOOL;			(* Program done. *)
	bBusy						:BOOL;			(* Program busy *)
	bError						:BOOL;			(* Error *)
	udnErrorNo					:UDINT;			(* Error number *)
	sErrorMsg					:STRING; 		(* Error message *)
END_VAR
VAR_IN_OUT
	(* Input Output variables / Ausgang Variablen *)
	Yaskawa					:ST_YASKAWA_REF;				(* The YASKAWA_REF data type  is an interface between the PLC and the YASKAWA and contains axis information *)
END_VAR
VAR
	(* Enummerations *)

	(* Variables *)

	(* References *)

	(* Interfaces *)

	(* Instances *)
	rtExecute						:R_TRIG;
	rtExtReset					:R_TRIG;
	rtDrivesOn					:R_TRIG;

END_VAR


rtExecute(CLK := bExecute
			      AND Yaskawa.stYaskawaToPlc.bAlarmErrorOccured);
rtDrivesOn(CLK := Yaskawa.stYaskawaToPlc.bServoIsOn
	   		        AND Yaskawa.stPlcToYaskawa.bExternalServoOn);

IF rtExecute.Q
     OR (rtDrivesOn.Q
	    AND Yaskawa.stYaskawaToPlc.bAlarmErrorOccured)
THEN
	bBusy := TRUE;
	Yaskawa.stPlcToYaskawa.bAlarmReset := TRUE;

ELSIF Yaskawa.stPlcToYaskawa.bAlarmReset
	   AND NOT Yaskawa.stYaskawaToPlc.bAlarmErrorOccured
THEN
	bBusy := FALSE;
	Yaskawa.stPlcToYaskawa.bAlarmReset := FALSE;
END_IF;

bDone := bExecute
		AND NOT bBusy
		AND NOT Yaskawa.stYaskawaToPlc.bAlarmErrorOccured;        (* Error *)

END_FUNCTION_BLOCK

// ---- POUs/Tc3 Objects/ExternalHardware/YASKAWA/FB_YASKAWA_StartPrg_1.TcPOU
FUNCTION_BLOCK FB_YASKAWA_StartPrg_1
(*

The function block used to start kuka

Constructor: 		Patryk Panylo
Company:		E. Riexinger GmbH
Date:			18.11.2016
Version:			1.00

Date:			Revision:		Who:				Comment

*)
VAR_INPUT
	(* Input variables / Eingang Variablen *)
	bEnable						:BOOL;			(* Signal FB enable *)
	bReset						:BOOL;			(* Signal reset *)
	bAutoHand					:BOOL;			(* Auto := TRUE, Hand := FALSE *)
	bStart						:BOOL;			(* Start program *)
	bStop						:BOOL;			(* Stop program *)
	nPrgNo						:INT;			(* Program number *)
END_VAR
VAR_OUTPUT
	(* Output variables / Ausgang Variablen *)
	bRunning					:BOOL;						(* Program running *)
	bDone						:BOOL;						(* Program done *)
	bBusy						:BOOL;						(* Program busy *)
	bError						:BOOL;						(* Error *)
	udnErrorNo					:UDINT;
END_VAR
VAR_IN_OUT
	(* Input Output variables / Ausgang Variablen *)
	Yaskawa					:ST_YASKAWA_REF;				(* The YASKAWA_REF data type  is an interface between the PLC and the YASKAWA and contains axis information *)
END_VAR
VAR
	(* Enummerations *)
	etYaskawaStart				:ET_YaskawaStart;

	(* Variables *)
	bFirstTime					:BOOL;

	nWatchdog					:INT;

	(* References *)

	(* Interfaces *)

	(* Instances *)
	rtStart						:R_TRIG;
	rtStop						:R_TRIG;
	rtReset						:R_TRIG;
	tonWatchdog					:TON;

END_VAR


IF NOT bEnable
THEN
	bDone := FALSE;					(* Program done *)
	bBusy := FALSE;                                  	(* Program not busy *)
	bError := FALSE;                                 	(* Program not error *)
	udnErrorNo := 0;                                 		(* Error number *)

	Yaskawa.stPlcToYaskawa.bCallMasterJob := FALSE;
	Yaskawa.stPlcToYaskawa.bExternalStart := FALSE;
	Yaskawa.stPlcToYaskawa.bExternalHold := FALSE;

	RETURN;
END_IF;

IF NOT bFirstTime
THEN
	tonWatchdog(IN := FALSE);

	Yaskawa.stPlcToYaskawa.bCallMasterJob := FALSE;
	Yaskawa.stPlcToYaskawa.bExternalStart := FALSE;
	Yaskawa.stPlcToYaskawa.bExternalHold := FALSE;

	etYaskawaStart := ET_YaskawaStart_eWaitExecute;              (* Next step *)

	bFirstTime := TRUE;
END_IF

rtReset(CLK := bReset);

IF rtReset.Q
     AND bError
THEN
	bError := FALSE;

	tonWatchdog(IN := FALSE);

	Yaskawa.stPlcToYaskawa.bCallMasterJob := FALSE;
	Yaskawa.stPlcToYaskawa.bExternalStart := FALSE;
	Yaskawa.stPlcToYaskawa.bExternalHold := FALSE;

	etYaskawaStart := ET_YaskawaStart_eWaitExecute;              (* Next step *)
END_IF

(* Wait for triger *)
rtStart(
	CLK := bStart
);

IF rtStart.Q
     AND Yaskawa.stYaskawaToPlc.bServoIsOn
     AND NOT Yaskawa.stYaskawaToPlc.bAlarmErrorOccured
THEN
	Yaskawa.stPlcToYaskawa.bCallMasterJob := FALSE;
	Yaskawa.stPlcToYaskawa.bExternalStart := FALSE;
	Yaskawa.stPlcToYaskawa.bExternalHold := FALSE;

	etYaskawaStart := ET_YaskawaStart_eWaitExecute;              (* Next step *)

END_IF

rtStop(
	CLK := bStop
);

IF rtStop.Q
     OR Yaskawa.stYaskawaToPlc.bAlarmErrorOccured
THEN
	Yaskawa.stPlcToYaskawa.bCallMasterJob := FALSE;
	Yaskawa.stPlcToYaskawa.bExternalStart := FALSE;
	Yaskawa.stPlcToYaskawa.bExternalHold := Yaskawa.stYaskawaToPlc.bOperatingRunning
										     AND NOT Yaskawa.stYaskawaToPlc.bAlarmErrorOccured;

	etYaskawaStart := ET_YaskawaStart_eWaitExecute;              (* Next step *)

END_IF

bRunning := Yaskawa.stYaskawaToPlc.bOperatingRunning;
Yaskawa.stPlcToYaskawa.nPrgNo := nPrgNo;

(* Send command *)
CASE etYaskawaStart OF

	ET_YaskawaStart_eWaitExecute:
		bBusy := FALSE;                                     	(* Program not busy *)
		bError := FALSE;                         		(* Program not error *)
		udnErrorNo := 0;                         		(* Error number *)

		IF rtStart.Q
     		     AND bAutoHand			(* Automatic *)
		     AND NOT bStop
		THEN
			nWatchdog := 0;
			bDone:= FALSE;                               		(* Program done *)
			bBusy := TRUE;                                  	(* Program busy *)

			tonWatchdog(IN := FALSE);

			Yaskawa.stPlcToYaskawa.bCallMasterJob := FALSE;
			Yaskawa.stPlcToYaskawa.bExternalStart := FALSE;
			Yaskawa.stPlcToYaskawa.bExternalHold := FALSE;

			IF Yaskawa.stYaskawaToPlc.bHold
			THEN
				etYaskawaStart := ET_YaskawaStart_eExternalStart;              (* Next step *)
			ELSE
				etYaskawaStart := ET_YaskawaStart_eCallMasterJob;              (* Next step *)
			END_IF
		END_IF

	ET_YaskawaStart_eCallMasterJob:
		nWatchdog := nWatchdog + 1;

		Yaskawa.stPlcToYaskawa.bCallMasterJob := TRUE;

		IF Yaskawa.stYaskawaToPlc.bTopMasterJob
		     AND Yaskawa.stYaskawaToPlc.bServoIsOn
		     AND NOT Yaskawa.stYaskawaToPlc.bAlarmErrorOccured
		THEN
			nWatchdog := 0;

			Yaskawa.stPlcToYaskawa.bCallMasterJob := FALSE;

			etYaskawaStart := ET_YaskawaStart_eExternalStart;              (* Next step *)

		ELSIF Yaskawa.stYaskawaToPlc.bAlarmErrorOccured
			    OR nWatchdog > 1000
		THEN
			Yaskawa.stPlcToYaskawa.bCallMasterJob := FALSE;
			
			udnErrorNo := 1;                     (* Error number *)
			
			etYaskawaStart := ET_YaskawaStart_eError;              (* Next step *)

		END_IF

	ET_YaskawaStart_eExternalStart:
		nWatchdog := nWatchdog + 1;

		Yaskawa.stPlcToYaskawa.bExternalStart := TRUE;

		IF Yaskawa.stYaskawaToPlc.bOperatingRunning
		     AND Yaskawa.stYaskawaToPlc.bServoIsOn
		     AND NOT Yaskawa.stYaskawaToPlc.bPrgDone
		     AND NOT Yaskawa.stYaskawaToPlc.bAlarmErrorOccured
		THEN
			nWatchdog := 0;

			Yaskawa.stPlcToYaskawa.bExternalStart := FALSE;

			etYaskawaStart := ET_YaskawaStart_eWfPrgDone;              (* Next step *)

		ELSIF Yaskawa.stYaskawaToPlc.bAlarmErrorOccured
			    OR nWatchdog > 1000
		THEN
			Yaskawa.stPlcToYaskawa.bExternalStart := FALSE;
			
			udnErrorNo := 2;                     (* Error number *)

			etYaskawaStart := ET_YaskawaStart_eError;              (* Next step *)

		END_IF

	ET_YaskawaStart_eWfPrgDone:
		IF (Yaskawa.stYaskawaToPlc.bInHome
		     OR Yaskawa.stYaskawaToPlc.bNotInCrashAreaMachine)
		    AND Yaskawa.stYaskawaToPlc.bPrgDone
	     	    AND NOT Yaskawa.stYaskawaToPlc.bAlarmErrorOccured
		THEN
			Yaskawa.stPlcToYaskawa.bCallMasterJob := FALSE;;
			Yaskawa.stPlcToYaskawa.bExternalStart := FALSE;

			etYaskawaStart := ET_YaskawaStart_eDone;              (* Next step *)

		ELSIF Yaskawa.stYaskawaToPlc.bAlarmErrorOccured
		THEN
			Yaskawa.stPlcToYaskawa.bCallMasterJob := FALSE;;
			Yaskawa.stPlcToYaskawa.bExternalStart := FALSE;

			udnErrorNo := 3;                     (* Error number *)

			etYaskawaStart := ET_YaskawaStart_eError;              (* Next step *)

		END_IF

	ET_YaskawaStart_eError:
		bBusy := FALSE;						(* Command busy *)
		bError := TRUE;						(* Command error  *)

		etYaskawaStart := ET_YaskawaStart_eNoExecute;

	ET_YaskawaStart_eDone:
		bDone := TRUE;						(* Command done *)
		bBusy := FALSE;						(* Command busy *)

		etYaskawaStart := ET_YaskawaStart_eNoExecute;

	ET_YaskawaStart_eNoExecute:
		IF NOT bStart
		THEN
			(* Reset outputs *)
			bDone := FALSE;						(* Command done *)
			bBusy := FALSE;						(* Command busy *)
			bError := FALSE;						(* Command error  *)

			nWatchdog := 0;

			etYaskawaStart := ET_YaskawaStart_eWaitExecute;
		END_IF
END_CASE;

END_FUNCTION_BLOCK

// ---- POUs/Tc3 Objects/File/CSV/FB_FileCSVHandler.TcPOU
FUNCTION_BLOCK FB_FileCSVHandler
(*

This function block is used to read and write datas into/from csv file.
None of the field value is containing any non-printing control characters like line feed, carriage return, quotation marks, semicolon... 

Constructor: 		Patryk Panylo
Company:			E. Riexinger GmbH
Date:				05.04.2019
Version:			1.00

Date:			Revision:		Who:				Comment
dd.mm.yyyy		x.xx			Initials			comment

*)

VAR_INPUT
	bEnable						:BOOL := FALSE;				(* Enable FB *)
	sNetID						:T_AmsNetID	:= '';			(* TwinCAT Net ID *)
	bExecute					:BOOL := FALSE;				(* Execute operation *)
	sFilePath					:T_MaxString := '';			(* File path *)
	sFileName					:T_MaxString := '';			(* File name *)
	bCommaSeparator				:BOOL := FALSE;				(* Enable comma csv separator *)
	dwOpenMode					:DWORD;				(*
															FOPEN_MODEREAD (16#0001)	"r": Opens for reading. If the file does not exist or cannot be found, the call fails.
															FOPEN_MODEWRITE (16#0002) "w": Opens an empty file for writing. If the given file exists, its contents are destroyed.
															FOPEN_MODEAPPEND (16#0004) "a": Opens for writing at the end of the file (appending) without removing the EOF marker before writing new data to the file; creates the file first if it doesn’t exist.
															FOPEN_MODEREAD OR FOPEN_MODEPLUS (16#0008) "r+": Opens for reading and writing. The file must exist.
															FOPEN_MODEWRITE OR FOPEN_MODEPLUS (16#0008) "w+": Opens an empty file for both reading and writing. If the given file exists, its contents are destroyed.
															FOPEN_MODEAPPEND OR FOPEN_MODEPLUS (16#0008)	 "a+": Opens for reading and appending; the appending operation includes the removal of the EOF marker before new data is written to the file and the EOF marker is restored after writing is complete; creates the file first if it doesn’t exist.
															When a file is opened with the "a" or "a+" access type, all write operations occur at the end of the file. The file pointer can be repositioned using FB_FileSeek, but is always moved back to the end of the file before any write operation is carried out. Thus, existing data cannot be overwritten.
															
															FOPEN_MODEBINARY (16#0010) "b": Open in binary (untranslated) mode.
															FOPEN_MODETEXT (16#0020) "t": Open in text (translated) mode.
														*)
	arsWriteRecords				:ARRAY[0..GVL_CSV.MAX_CSV_ROWS, 0..GVL_CSV.MAX_CSV_COLUMNS ] OF STRING(GVL_CSV.MAX_CSV_FIELD_LENGTH);			(* Write records *)
	udnRowUsingMax				:UDINT;						(* Maximal number of using rows *)
	udnColumnUsingMax			:UDINT;						(* Maximal number of using columns *)																				
	tTimeout					:TIME := T#1S;				(* States the time before the function is cancelled *)
END_VAR
VAR_OUTPUT
	arsReadRecords				:ARRAY[0..GVL_CSV.MAX_CSV_ROWS, 0..GVL_CSV.MAX_CSV_COLUMNS ] OF STRING(GVL_CSV.MAX_CSV_FIELD_LENGTH);			(* Read records *)																										
	bBusy						:BOOL;					(* Program busy *)
	bDone						:BOOL;					(* Program done *)
	bError						:BOOL;					(* Program error *)
	udnErrNo					:UDINT;					(* Error number *)
END_VAR
VAR_IN_OUT

END_VAR
VAR
	(* Enummerations *)
	etCSVState					:ET_CSV_State := ET_CSV_State_eWaitExecute;
	
	(* Variables *)
	bFirstTime					:BOOL;					(* First PLC cycle *)

	dwModeCache					:DWORD;					(* Contains the mode in which the file is to be opened *)
	sPathName					:STRING;				(* Contains the path and filename for the file to be opened *)
	hFileHandle					:UINT;					(* File handle *)

	udnWriteCounter				:UDINT;
	udnReadCounter				:UDINT;

	udnRowCounter				:UDINT;
	udnColumnCounter			:UDINT;
	
	sCSVLine					:T_MaxString := '';		(* Single CSV text line (row, record), we are using string as record buffer (your are able to see created fields) *)
	sCSVField					:T_MaxString := '';		(* Single CSV field value (column, record field) *)
	
	(* Instances *)
	fbCreateDir					:FB_CreateDir;			(* Create direction *)
	
	fbFileOpen					:FB_FileOpen;			(* File open *)
	fbFileClose					:FB_FileClose;			(* File close *)

	fbFilePuts					:FB_FilePuts;			(* Writes one record (line) *)
	fbWriter					:FB_CSVMemBufferWriter;	(* Helper function block used to create CSV data bytes (single record line) *)
	
	fbFileGets					:FB_FileGets;			(* Reads one record (line) *)
	fbReader					:FB_CSVMemBufferReader;	(* Helper function block used to parse CSV data bytes (single record line) *)
END_VAR
VAR CONSTANT
	sFileSuffix					:STRING(5) := 'csv';
END_VAR

IF NOT bEnable				(* Enable FB *)
THEN
	bFirstTime := FALSE;		(* First PLC cycle *)
	bBusy := FALSE;			(* Program busy *)
	bDone := FALSE;			(* Program done *)
	bError := FALSE;			(* Program error *)
	udnErrNo := 0;				(* Error number *)
	RETURN;
END_IF

IF NOT bFirstTime
THEN
	IF bCommaSeparator
	THEN
		DEFAULT_CSV_FIELD_SEP := 16#2C;			(* Comma ASCII code *)
	ELSE
		DEFAULT_CSV_FIELD_SEP := 16#3B;			(* Semicolon ASCII code *)
	END_IF

	etCSVState := ET_CSV_State_eWaitExecute;

	bFirstTime := TRUE;
END_IF


(* Sequence state for open, read/write and close the file *)
CASE etCSVState
OF
	ET_CSV_State_eWaitExecute:
		IF bExecute
		THEN				
			fbCreateDir(
				sNetId:= sNetID,
				sPathName:= sFilePath,
				ePath:= PATH_GENERIC,
				bExecute := FALSE, 
				tTimeout:= tTimeout
			);
		
			fbFileOpen(								(* File open *)
				sNetId := sNetID,
				nMode := dwOpenMode, 
				ePath := PATH_GENERIC,
				bExecute := FALSE,
				tTimeout := tTimeout 
			);			
			fbFileClose(							(* File close *)
				sNetId := sNetID, 
				bExecute := FALSE,
				tTimeout := tTimeout 
			);			
			
			fbFilePuts(								(* Writes one record (line) *)
				sNetId := sNetID,
				bExecute := FALSE,
				tTimeout := tTimeout 
			);			

			fbFileGets(								(* Writes one record (line) *)
				sNetId := sNetID,
				bExecute := FALSE,
				tTimeout := tTimeout 
			);
	
			(* Create data path *)
			sPathName := CONCAT(sFilePath, CONCAT(sFileName, CONCAT('.', sFileSuffix)));
	
			IF sPathName <> ''
			   AND dwOpenMode <> 0
			THEN
				udnErrNo := 0;
			
				etCSVState := ET_CSV_State_eCreateDir;			(* Next step *)
	
			ELSE
				udnErrNo := 1;
	
				etCSVState := ET_CSV_State_eError;				(* Next step *)
	
			END_IF
				
			bBusy := TRUE;
			bDone := FALSE;
			bError := FALSE;
			hFileHandle := 0;
			udnRowCounter := 0;
			udnColumnCounter := 0;

		END_IF
		
	(* Create direction *)
	ET_CSV_State_eCreateDir:
		fbCreateDir(bExecute := FALSE);
		fbCreateDir(
			sPathName := sFilePath, 
			bExecute := TRUE
		);

		etCSVState := ET_CSV_State_eChkCreateDir;				(* Next step *)

	ET_CSV_State_eChkCreateDir:	
		fbCreateDir(bExecute := FALSE);
	
		IF NOT fbCreateDir.bBusy
		THEN
			IF NOT fbCreateDir.bError
			THEN
				etCSVState := ET_CSV_State_eFileOpen;				(* Next step *)
			ELSE
				IF  fbCreateDir.nErrId = 16#723 	(* 0x723 Folder is allready existing or invalid sPathName or ePath parameter.*)
				THEN
					etCSVState := ET_CSV_State_eFileOpen;				(* Next step *)
				ELSE
					udnErrNo := fbFilePuts.nErrId;	
				
					etCSVState := ET_CSV_State_eError;					(* Next step *)
				END_IF
			END_IF
		END_IF
				
	(* Open the file *)
	ET_CSV_State_eFileOpen:
		fbFileOpen(bExecute := FALSE);
		fbFileOpen(
			sPathName := sPathName, 
			bExecute := TRUE
		);

		etCSVState := ET_CSV_State_eChkFileOpen;				(* Next step *)

	(* Check open the file *)
	ET_CSV_State_eChkFileOpen:
		fbFileOpen(bExecute := FALSE);
		
		IF NOT fbFileOpen.bBusy
		THEN
			IF NOT fbFileOpen.bError
			THEN
				hFileHandle := fbFileOpen.hFile;

				(* Choose write or read datas *)
				IF fbFileOpen.nMode = (FOPEN_MODEWRITE OR FOPEN_MODETEXT)
				THEN
					etCSVState := ET_CSV_State_eConvertRecord;			(* Next step *)

				ELSIF fbFileOpen.nMode = (FOPEN_MODEAPPEND OR FOPEN_MODETEXT)
				THEN
					etCSVState := ET_CSV_State_eConvertRecord;			(* Next step *)

				ELSIF fbFileOpen.nMode = (FOPEN_MODEREAD OR FOPEN_MODETEXT)
				THEN
					etCSVState := ET_CSV_State_eFileGets;			(* Next step *)
				
				ELSE
					udnErrNo := 2;
	
					etCSVState := ET_CSV_State_eError;				(* Next step *)

				END_IF
			ELSE
				udnErrNo := fbFileOpen.nErrId;
	
				etCSVState := ET_CSV_State_eError;					(* Next step *)
				
			END_IF
		END_IF

	(* Convert one PLC record to CSV format *)		
	ET_CSV_State_eConvertRecord:
		sCSVLine := '';
		fbWriter.eCmd := eEnumCmd_First;			(* Write first field value *)
		
		IF udnRowCounter <= MIN(udnRowUsingMax, GVL_CSV.MAX_CSV_ROWS) 
		THEN	
			FOR udnColumnCounter := 0 TO MIN(udnColumnUsingMax, GVL_CSV.MAX_CSV_COLUMNS) BY 1 
			DO	
				(* Get field value *)	
				sCSVField := STRING_TO_CSVFIELD(			
								arsWriteRecords[udnRowCounter, udnColumnCounter], 
								FALSE
							 );
		
				(* Add new field to the record buffer *)
				fbWriter(
					pBuffer := ADR(sCSVLine), 
					cbBuffer := SIZEOF(sCSVLine) - 1, 
					putValue := sCSVField, 
					pValue := 0, 
					cbValue := 0,
					bCRLF := (udnColumnCounter = MIN(udnColumnUsingMax, GVL_CSV.MAX_CSV_COLUMNS))			(* bCRLF == TRUE => Write CRLF after the last field value *)
				);
				
				IF fbWriter.bOk 
				THEN
					fbWriter.eCmd := eEnumCmd_Next;			(* Write next field value *)
					
				ELSE(* Error *)
					udnErrNo := 3;	
				
					etCSVState := ET_CSV_State_eError;					(* Next step *)
					
					RETURN;
				END_IF
		
			END_FOR
		
			(* FB_FilePuts adds allready CR (carriage return) to the written line.
			   We have to replace the $R$L characters with $L character to avoid double CR. *)
			IF RIGHT(sCSVLine, 2) = '$R$L' 
			THEN
				sCSVLine := REPLACE(sCSVLine, '$L', 2, LEN(sCSVLine) - 1);
			END_IF
		
			udnRowCounter := udnRowCounter + 1;					(* Increment number of created records (rows) *)
			
			etCSVState := ET_CSV_State_eFilePuts;				(* Write record to the file *)
		
		ELSE			(* All rows written => Close file *)
			udnWriteCounter := udnWriteCounter + 1;	
		
			etCSVState := ET_CSV_State_eFileClose;
		END_IF
		
		
	(* Writes one record (line) *)
	ET_CSV_State_eFilePuts:
		fbFilePuts(bExecute := FALSE);
		
		fbFilePuts(	
			hFile := hFileHandle, 
			sLine := sCSVLine, 
			bExecute := TRUE
		);

		etCSVState := ET_CSV_State_eChkFilePuts;				(* Next step *)

	(* Check write the file *)
	ET_CSV_State_eChkFilePuts:
		fbFilePuts(bExecute := FALSE);
		
		IF NOT fbFilePuts.bBusy
		THEN
			IF NOT fbFilePuts.bError
			THEN			
				etCSVState := ET_CSV_State_eConvertRecord;					(* Next step *)
				
			ELSE
				udnErrNo := fbFilePuts.nErrId;
	
				etCSVState := ET_CSV_State_eError;					(* Next step *)
				
			END_IF
		END_IF

	(* Read single line (record) *)
	ET_CSV_State_eFileGets:
		fbFileGets(bExecute := FALSE);
		
		fbFileGets(	
			hFile := hFileHandle, 
			bExecute := TRUE
		);

		etCSVState := ET_CSV_State_eChkFileGets;				(* Next step *)

	(* Check read the file *)
	ET_CSV_State_eChkFileGets:
		fbFileGets(bExecute := FALSE);
		
		sCSVLine := fbFileGets.sLine;
		
		IF NOT fbFileGets.bBusy
		THEN
			IF NOT fbFileGets.bError
			THEN				
				IF fbFileGets.bEOF 
				THEN
					udnReadCounter := udnReadCounter + 1;
				
					etCSVState := ET_CSV_State_eFileClose;			(* End of file reached => Close source file *)
				ELSE
					(* FB_FileGets returns text line without the CR (carriage return) character.
					   We have to restore the CR character (replace the $L character with $R$L characters) *)
					IF RIGHT(sCSVLine, 1) = '$L' 
					THEN
						sCSVLine := REPLACE(sCSVLine, '$R$L', 2, LEN(sCSVLine));
					END_IF

					etCSVState := ET_CSV_State_eParseSingleRecord;
					
				END_IF
				
			ELSE
				udnErrNo := fbFilePuts.nErrId;
	
				etCSVState := ET_CSV_State_eError;					(* Next step *)
				
			END_IF
		END_IF
		
	(* Parse single record *)
	ET_CSV_State_eParseSingleRecord:
		fbReader.eCmd := eEnumCmd_First;			(* Read first field value *)
		
		REPEAT
			fbReader(
				pBuffer := ADR(sCSVLine), 
				cbBuffer := SIZEOF(sCSVLine), 
				getValue => sCSVField
			);
			
			IF fbReader.bOk THEN
				fbReader.eCmd := eEnumCmd_Next;			(* Read next field value *)

				IF udnRowCounter <= MIN(udnRowUsingMax, GVL_CSV.MAX_CSV_ROWS) 
				THEN
					IF udnColumnCounter <= MIN(udnColumnUsingMax, GVL_CSV.MAX_CSV_COLUMNS) 
					THEN
						(* Save or use the field value *)
						arsReadRecords[udnRowCounter, udnColumnCounter] := CSVFIELD_TO_STRING(sCSVField, FALSE);
					END_IF
				END_IF

				udnColumnCounter := udnColumnCounter + 1;			(* Increment number of read columns *)
				
				IF fbReader.bCRLF			(* CRLF == TRUE => End of reacord reached *)
				THEN
					udnRowCounter := udnRowCounter + 1;				(* Increment number of read records *)
					udnColumnCounter := 0;			(* Reset number of columns *)
				END_IF

			ELSE			(* Error: End of record reached or all fields read *)
				etCSVState := ET_CSV_State_eFileGets;(* Try to read next line *)
				
			END_IF
			
		UNTIL NOT fbReader.bOk		
		END_REPEAT
				
	(* Close the file *)
	ET_CSV_State_eFileClose:
		fbFileClose(bExecute := FALSE);
		
		fbFileClose(	
			hFile := hFileHandle, 
			bExecute := TRUE
		);

		etCSVState := ET_CSV_State_eChkFileClose;				(* Next step *)

	(* Check close the file *)
	ET_CSV_State_eChkFileClose:
		fbFileClose(bExecute := FALSE);
	
		IF NOT fbFileClose.bBusy
		THEN
			hFileHandle := 0;
		
			IF NOT fbFileClose.bError
			THEN
				etCSVState := ET_CSV_State_eDone;					(* Next step *)

			ELSE
				udnErrNo := fbFileClose.nErrId;
	
				etCSVState := ET_CSV_State_eError;					(* Next step *)
				
			END_IF
		END_IF

	ET_CSV_State_eDone:
		bBusy := FALSE;
		bDone := TRUE;
		bError := FALSE;
		
		etCSVState := ET_CSV_State_eNoExecute;					(* Next step *)

	ET_CSV_State_eError:
		IF hFileHandle <> 0
		THEN
			bDone := FALSE;
			bError := TRUE;
			
			etCSVState := ET_CSV_State_eFileClose;					(* Next step *)

		ELSE
			bBusy := FALSE;
			bDone := FALSE;
			bError := TRUE;
	
			etCSVState := ET_CSV_State_eNoExecute;					(* Next step *)
		END_IF

	ET_CSV_State_eNoExecute:
		IF NOT bExecute
		THEN
			bBusy := FALSE;
			bDone := FALSE;
			bError := FALSE;

			etCSVState := ET_CSV_State_eWaitExecute;			(* Next step *)

		END_IF

END_CASE

END_FUNCTION_BLOCK

// ---- POUs/Tc3 Objects/File/TXT/FB_FileHandlerBinary_1.TcPOU
FUNCTION_BLOCK FB_FileHandlerBinary_1
(*

This function block is used to read and write binary datas in/from file.

Constructor: 		Patryk Panylo
Company:		E. Riexinger GmbH
Date:			10.06.2013
Version:			1.00

Date:			Revision:		Who:				Comment
dd.mm.yyyy		x.xx			Initials			comment

*)

VAR_INPUT
	bEnable						:BOOL;					(* Enable FB *)
	bExecute					:BOOL;					(* Execute operation *)
	sFilePath					:STRING;				(* File path *)
	sFileName					:STRING;				(* File name *)
	sFileSuffix					:STRING := 'dat';			(* Suffix of file *)
	bFileWrite					:BOOL;					(* Write file *)
	bFileRead					:BOOL;					(* Read file *)
	dwDataBuffer					:POINTER TO DWORD;				(* Contains the address of the buffer containing the data to be read/written ADR *)
	udnDataBufLen				:UDINT;					(* Contains the number of bytes to be written SIZEOF *)
	tTimeout						:TIME := t#1s;				(* States the time before the function is cancelled *)
END_VAR
VAR_OUTPUT
	bBusy						:BOOL;					(* Program busy *)
	bDone						:BOOL;					(* Program done *)
	bError						:BOOL;					(* Program error *)
	udnErrNo					:UDINT;					(* Error number *)
END_VAR
VAR_IN_OUT

END_VAR
VAR
	(* Enummerations *)
	enStep						: (eWaitExecute := 0, eChkFileName,  eChkBufLen, eFileOpen, eChkFileOpen, eFileWrite, eChkFileWrite, eFileRead, eChkFileRead, eFileClose, eChkFileClose, eDone, eError, eNotExecute);			(* Sequence state for open, read/write and close the file *)

	(* Variables *)
	bFirstTime					:BOOL;					(* First PLC cycle *)

	dwMode						:DWORD;				(* Contains the mode in which the file is to be opened *)
	sPathName					:STRING;				(* Contains the path and filename for the file to be opened *)
	hFileHandle					:UINT;					(* File handle *)

	unWriteCounter				:UINT;
	unReadCounter				:UINT;

	(* Instances *)
	fbFileOpen					:FB_FileOpen;			(* File open *)
	fbFileClose					:FB_FileClose;			(* File close *)
	fbFileRead					:FB_FileRead;			(* File read *)
	fbFileWrite					:FB_FileWrite;				(* File write *)

END_VAR

IF NOT bEnable				(* Enable FB *)
THEN
	bFirstTime := FALSE;		(* First PLC cycle *)
	bBusy := FALSE;			(* Program busy *)
	bDone := FALSE;			(* Program done *)
	bError := FALSE;			(* Program error *)
	udnErrNo := 0;				(* Error number *)
	RETURN;
END_IF

IF NOT bFirstTime
THEN
	enStep := eWaitExecute;

	bFirstTime := TRUE;
END_IF


(* Sequence state for open, read/write and close the file *)
CASE enStep
OF

	eWaitExecute:
		IF bExecute
		THEN
			fbFileOpen.bExecute := FALSE;			(* File open *)
			fbFileClose.bExecute := FALSE;			(* File close *)
			fbFileRead.bExecute := FALSE;			(* File read *)
			fbFileWrite.bExecute := FALSE;			(* File write *)

			bDone := FALSE;
			bError := FALSE;
			udnErrNo := 0;

			IF bFileWrite
			THEN
				dwMode := FOPEN_MODEWRITE OR FOPEN_MODEBINARY;

				enStep := eChkFileName;			(* Next step *)

			ELSIF bFileRead
			THEN
				dwMode := FOPEN_MODEREAD OR FOPEN_MODEBINARY;

				enStep := eChkFileName;			(* Next step *)

			ELSE
				RETURN;
			END_IF

			bBusy := TRUE;

		END_IF

	(* Check file name and path *)
	eChkFileName:

		sPathName := CONCAT(
						sFilePath, CONCAT(
									sFileName, CONCAT(
												'.', sFileSuffix)));

		IF sFilePath <> ''
		     AND sFileName <> ''
		     AND sFileSuffix <> ''
		THEN
			enStep := eChkBufLen;			(* Next step *)

		ELSE
			udnErrNo := INT_TO_UINT(eChkFileName);

			enStep := eError;				(* Next step *)

		END_IF


	(* Check buffer lenght *)
	eChkBufLen:
		IF udnDataBufLen = 0
		THEN
			enStep := eDone;				(* Next step *)
	
		ELSE
			enStep := eFileOpen;			(* Next step *)
		
		END_IF

	(* Open the file *)
	eFileOpen:
		fbFileOpen.bExecute := TRUE;

		enStep := eChkFileOpen;				(* Next step *)

	(* Check open the file *)
	eChkFileOpen:
		IF NOT fbFileOpen.bBusy
		THEN
			IF NOT fbFileOpen.bError
			THEN
				fbFileOpen.bExecute := FALSE;
				hFileHandle := fbFileOpen.hFile;

				(* Choose write or read datas *)
				IF fbFileOpen.nMode = (FOPEN_MODEWRITE OR FOPEN_MODEBINARY)
				THEN
					enStep := eFileWrite;			(* Next step *)
	
				ELSIF fbFileOpen.nMode = (FOPEN_MODEREAD OR FOPEN_MODEBINARY)
				THEN
					enStep := eFileRead;			(* Next step *)

				ELSE
					enStep := eFileClose;			(* Next step *)
	
				END_IF

			ELSE
				fbFileOpen.bExecute := FALSE;
				udnErrNo := fbFileOpen.nErrId;
	
				enStep := eError;					(* Next step *)
				
			END_IF
		END_IF

	(* Write the file *)
	eFileWrite:
		fbFileWrite.bExecute := TRUE;

		enStep := eChkFileWrite;				(* Next step *)

	(* Check write the file *)
	eChkFileWrite:
		IF NOT fbFileWrite.bBusy
		THEN
			IF fbFileRead.cbRead = 0
				AND NOT fbFileRead.bError
			THEN
				fbFileWrite.bExecute := FALSE;
				unWriteCounter := 0;
	
				enStep := eFileClose;				(* Next step *)	
				
			ELSIF (fbFileWrite.cbWrite >= SIZEOF(dwDataBuffer))
			    AND NOT fbFileWrite.bError
			THEN
				fbFileWrite.bExecute := FALSE;
				unWriteCounter := unWriteCounter + 1;

				enStep := eFileClose;				(* Next step *)

			ELSIF  fbFileWrite.bError
			THEN
				fbFileWrite.bExecute := FALSE;
				udnErrNo := fbFileWrite.nErrId;

				enStep := eError;					(* Next step *)
				
			END_IF
		END_IF

	(* Read the file *)
	eFileRead:
		fbFileRead.bExecute := TRUE;

		enStep := eChkFileRead;				(* Next step *)

	(* Check read the file *)
	eChkFileRead:
		IF NOT fbFileRead.bBusy
		THEN
			IF fbFileRead.cbRead = 0
				AND NOT fbFileRead.bError
			THEN
				fbFileRead.bExecute := FALSE;
				unReadCounter := 0;
	
				enStep := eFileClose;				(* Next step *)	
				
			ELSIF (fbFileRead.cbRead >= SIZEOF(dwDataBuffer))
			     AND NOT fbFileRead.bError
			THEN
				fbFileRead.bExecute := FALSE;
				unReadCounter := unReadCounter + 1;
	
				enStep := eFileClose;				(* Next step *)

			ELSIF  fbFileRead.bError
			THEN
				fbFileRead.bExecute := FALSE;
				udnErrNo := fbFileRead.nErrId;
	
				enStep := eError;					(* Next step *)
				
			END_IF
		END_IF

	(* Close the file *)
	eFileClose:
		fbFileClose.bExecute := TRUE;

		enStep := eChkFileClose;				(* Next step *)

	(* Check close the file *)
	eChkFileClose:
		IF NOT fbFileClose.bBusy
		THEN
			IF NOT fbFileClose.bError
			THEN
				fbFileClose.bExecute := FALSE;
				enStep := eDone;					(* Next step *)

				IF bError
				THEN
					enStep := eError;				(* Next step *)
				END_IF

			ELSE
				fbFileClose.bExecute := FALSE;
				udnErrNo := fbFileClose.nErrId;
	
				enStep := eError;					(* Next step *)
				
			END_IF
		END_IF

	eDone:
		bBusy := FALSE;
		bDone := TRUE;
		bError := FALSE;
		udnErrNo := 0;

		enStep := eNotExecute;					(* Next step *)

	eError:
		IF NOT bError
		     AND hFileHandle <> 0
		THEN
			bDone := FALSE;
			bError := TRUE;

			enStep := eFileClose;					(* Next step *)

		ELSE
			bBusy := FALSE;
			bDone := FALSE;
			bError := TRUE;
	
			enStep := eNotExecute;					(* Next step *)
		END_IF

	eNotExecute:
		IF NOT bExecute
		THEN
			bBusy := FALSE;
			bDone := FALSE;
			bError := FALSE;
			udnErrNo := 0;

			enStep := eWaitExecute;			(* Next step *)

		END_IF

END_CASE


fbFileOpen(
	sNetId := '',
	sPathName := sPathName,
	nMode := dwMode,
	ePath := PATH_GENERIC,
	tTimeout := tTimeout);
fbFileClose(
	sNetId := '',
	hFile := hFileHandle,
	tTimeout := tTimeout );
fbFileWrite(
	sNetId := '',
	hFile := hFileHandle,
	pWriteBuff := dwDataBuffer,
	cbWriteLen := udnDataBufLen,
	tTimeout := tTimeout);
fbFileRead(
	sNetId := '',
	hFile := hFileHandle,
	pReadBuff := dwDataBuffer,
	cbReadLen := udnDataBufLen,
	tTimeout := tTimeout);

END_FUNCTION_BLOCK

// ---- POUs/Tc3 Objects/File/TXT/FB_FileHandler_1.TcPOU
FUNCTION_BLOCK FB_FileHandler_1
(*

This function block is used to read and write binary datas in/from file.

Constructor: 		Patryk Panylo
Company:		E. Riexinger GmbH
Date:			10.06.2013
Version:			1.00

Date:			Revision:		Who:				Comment
dd.mm.yyyy		x.xx			Initials			comment

*)

VAR_INPUT
	bEnable						:BOOL;					(* Enable FB *)
	bExecute					:BOOL;					(* Execute operation *)
	sFilePath					:STRING;				(* File path *)
	sFileName					:STRING;				(* File name *)
	sFileSuffix					:STRING := 'dat';			(* Suffix of file *)
	dwOpenMode				:DWORD;				(*
															FOPEN_MODEREAD (16#0001)	"r": Opens for reading. If the file does not exist or cannot be found, the call fails.
															FOPEN_MODEWRITE (16#0002) "w": Opens an empty file for writing. If the given file exists, its contents are destroyed.
															FOPEN_MODEAPPEND (16#0004) "a": Opens for writing at the end of the file (appending) without removing the EOF marker before writing new data to the file; creates the file first if it doesn’t exist.
															FOPEN_MODEREAD OR FOPEN_MODEPLUS (16#0008) "r+": Opens for reading and writing. The file must exist.
															FOPEN_MODEWRITE OR FOPEN_MODEPLUS (16#0008) "w+": Opens an empty file for both reading and writing. If the given file exists, its contents are destroyed.
															FOPEN_MODEAPPEND OR FOPEN_MODEPLUS (16#0008)	 "a+": Opens for reading and appending; the appending operation includes the removal of the EOF marker before new data is written to the file and the EOF marker is restored after writing is complete; creates the file first if it doesn’t exist.
															When a file is opened with the "a" or "a+" access type, all write operations occur at the end of the file. The file pointer can be repositioned using FB_FileSeek, but is always moved back to the end of the file before any write operation is carried out. Thus, existing data cannot be overwritten.
															
															FOPEN_MODEBINARY (16#0010) "b": Open in binary (untranslated) mode.
															FOPEN_MODETEXT (16#0020) "t": Open in text (translated) mode.
														*)
	sWriteRecord					:T_MaxString;				(* Record to write *)
	tTimeout						:TIME := t#1s;				(* States the time before the function is cancelled *)
END_VAR
VAR_OUTPUT
	sReadRecord				:T_MaxString;				(* Record to read *)
	bBusy						:BOOL;					(* Program busy *)
	bDone						:BOOL;					(* Program done *)
	bError						:BOOL;					(* Program error *)
	udnErrNo					:UDINT;					(* Error number *)
END_VAR
VAR_IN_OUT

END_VAR
VAR
	(* Enummerations *)
	enStep						: (eWaitExecute := 0, eChkFileName,  eChkBufLen, eCreateDir, eChkCreateDir, eFileOpen, eChkFileOpen, eFileWrite, eChkFileWrite, eFileRead, eChkFileRead, eFileClose, eChkFileClose, eDone, eError, eNotExecute);			(* Sequence state for open, read/write and close the file *)

	(* Variables *)
	bFirstTime					:BOOL;					(* First PLC cycle *)

	dwModeCache				:DWORD;				(* Contains the mode in which the file is to be opened *)
	sWriteRecordCache			:T_MaxString;				(* Record to write *)
	sPathName					:STRING;				(* Contains the path and filename for the file to be opened *)
	hFileHandle					:UINT;					(* File handle *)

	unWriteCounter				:UINT;
	unReadCounter				:UINT;

	(* Instances *)
	fbCreateDir					:FB_CreateDir;			(* File open *)
	fbFileOpen					:FB_FileOpen;			(* File open *)
	fbFileClose					:FB_FileClose;			(* File close *)
	fbFileRead					:FB_FileRead;			(* File read *)
	fbFileWrite					:FB_FileWrite;				(* File write *)

END_VAR

IF NOT bEnable				(* Enable FB *)
THEN
	bFirstTime := FALSE;		(* First PLC cycle *)
	bBusy := FALSE;			(* Program busy *)
	bDone := FALSE;			(* Program done *)
	bError := FALSE;			(* Program error *)
	udnErrNo := 0;				(* Error number *)
	RETURN;
END_IF

IF NOT bFirstTime
THEN
	enStep := eWaitExecute;

	bFirstTime := TRUE;
END_IF


(* Sequence state for open, read/write and close the file *)
CASE enStep
OF

	eWaitExecute:
		IF bExecute
		THEN
			fbFileOpen.bExecute := FALSE;			(* File open *)
			fbFileClose.bExecute := FALSE;			(* File close *)
			fbFileRead.bExecute := FALSE;			(* File read *)
			fbFileWrite.bExecute := FALSE;			(* File write *)

			bDone := FALSE;
			bError := FALSE;
			udnErrNo := 0;

			sWriteRecordCache := sWriteRecord;

			IF dwOpenMode <> 0
			THEN
				dwModeCache := dwOpenMode;

				enStep := eChkFileName;			(* Next step *)

			ELSE
				RETURN;
			END_IF

			bBusy := TRUE;

		END_IF

	(* Check file name and path *)
	eChkFileName:

		sPathName := CONCAT(
						sFilePath, CONCAT(
									sFileName, CONCAT(
												'.', sFileSuffix)));

		IF sFilePath <> ''
		     AND sFileName <> ''
		     AND sFileSuffix <> ''
		THEN
			enStep := eChkBufLen;			(* Next step *)

		ELSE
			udnErrNo := INT_TO_UINT(eChkFileName);

			enStep := eError;				(* Next step *)

		END_IF


	(* Check buffer lenght *)
	eChkBufLen:
		IF LEN(sWriteRecordCache) = 0
		THEN
			enStep := eDone;				(* Next step *)
	
		ELSE
			(*enStep := eCreateDir;			(* Next step *)*)
			enStep := eFileOpen;			(* Next step *)
		END_IF

	(* Create direction *)
	eCreateDir:
		fbCreateDir.bExecute := TRUE;

		enStep := eChkCreateDir;				(* Next step *)

	eChkCreateDir:
		IF NOT fbCreateDir.bBusy
		THEN
			IF NOT fbCreateDir.bError
			THEN
				fbCreateDir.bExecute := FALSE;

				enStep := eFileOpen;				(* Next step *)
			ELSE
				fbCreateDir.bExecute := FALSE;

				IF  fbCreateDir.nErrId = 16#70C 	(* 0x70C Folder is allready existing or invalid sPathName or ePath parameter.*)
				THEN
					enStep := eFileOpen;				(* Next step *)
				ELSE
					enStep := eError;					(* Next step *)
				END_IF
			END_IF
		END_IF

	(* Open the file *)
	eFileOpen:
		IF LEN(sWriteRecordCache) > 254
		THEN
			sWriteRecordCache := DELETE(
								sWriteRecordCache,
								LEN(sWriteRecordCache) + 1 - 254, 254
							    );
		END_IF

		fbFileOpen.bExecute := TRUE;

		enStep := eChkFileOpen;				(* Next step *)

	(* Check open the file *)
	eChkFileOpen:
		IF NOT fbFileOpen.bBusy
		THEN
			IF NOT fbFileOpen.bError
			THEN
				fbFileOpen.bExecute := FALSE;
				hFileHandle := fbFileOpen.hFile;

				(* Choose write or read datas *)
				IF fbFileOpen.nMode = FOPEN_MODEWRITE
				THEN
				
					enStep := eFileWrite;			(* Next step *)

				ELSIF fbFileOpen.nMode = FOPEN_MODEAPPEND
				THEN
	
					enStep := eFileWrite;			(* Next step *)

				ELSIF fbFileOpen.nMode = FOPEN_MODEREAD
				THEN
					enStep := eFileRead;			(* Next step *)
				
				ELSE
					enStep := eFileClose;			(* Next step *)

				END_IF

			ELSE
				fbFileOpen.bExecute := FALSE;
				udnErrNo := fbFileOpen.nErrId;
	
				enStep := eError;					(* Next step *)
				
			END_IF
		END_IF

	(* Write the file *)
	eFileWrite:
		fbFileWrite.bExecute := TRUE;

		enStep := eChkFileWrite;				(* Next step *)

	(* Check write the file *)
	eChkFileWrite:
		IF NOT fbFileWrite.bBusy
		THEN
			IF fbFileWrite.cbWrite = 0
			    AND NOT fbFileWrite.bError
			THEN
				fbFileWrite.bExecute := FALSE;
				unWriteCounter := 0;

				enStep := eFileClose;				(* Next step *)
				
			ELSIF (fbFileWrite.cbWrite >= INT_TO_UDINT(LEN(sWriteRecordCache)))
			    AND NOT fbFileWrite.bError
			THEN
				fbFileWrite.bExecute := FALSE;
				unWriteCounter := unWriteCounter + 1;

				enStep := eFileClose;				(* Next step *)

			ELSIF  fbFileWrite.bError
			THEN
				fbFileWrite.bExecute := FALSE;
				udnErrNo := fbFileWrite.nErrId;

				enStep := eError;					(* Next step *)
				
			END_IF
		END_IF

	(* Read the file *)
	eFileRead:
		fbFileRead.bExecute := TRUE;

		enStep := eChkFileRead;				(* Next step *)

	(* Check read the file *)
	eChkFileRead:
		IF NOT fbFileRead.bBusy
		THEN
			IF fbFileRead.cbRead = 0
			     AND NOT fbFileRead.bError
			THEN
				fbFileRead.bExecute := FALSE;
				unReadCounter := 0;
	
				enStep := eFileClose;				(* Next step *)

			ELSIF (fbFileRead.cbRead >= INT_TO_UDINT(LEN(sReadRecord)))
			     AND NOT fbFileRead.bError
			THEN
				fbFileRead.bExecute := FALSE;
				unReadCounter := unReadCounter + 1;
	
				enStep := eFileClose;				(* Next step *)

			ELSIF fbFileRead.bEOF
			     AND NOT fbFileRead.bError
			THEN
				fbFileRead.bExecute := FALSE;
	
				enStep := eFileClose;				(* Next step *)
				
			ELSIF  fbFileRead.bError
			THEN
				fbFileRead.bExecute := FALSE;
				udnErrNo := fbFileRead.nErrId;
	
				enStep := eError;					(* Next step *)
				
			END_IF
		END_IF

	(* Close the file *)
	eFileClose:
		fbFileClose.bExecute := TRUE;

		enStep := eChkFileClose;				(* Next step *)

	(* Check close the file *)
	eChkFileClose:
		IF NOT fbFileClose.bBusy
		THEN
			IF NOT fbFileClose.bError
			THEN
				fbFileClose.bExecute := FALSE;
				enStep := eDone;					(* Next step *)

				IF bError
				THEN
					enStep := eError;				(* Next step *)
				END_IF

			ELSE
				fbFileClose.bExecute := FALSE;
				udnErrNo := fbFileClose.nErrId;
	
				enStep := eError;					(* Next step *)
				
			END_IF
		END_IF

	eDone:
		bBusy := FALSE;
		bDone := TRUE;
		bError := FALSE;
		udnErrNo := 0;

		enStep := eNotExecute;					(* Next step *)

	eError:
		IF NOT bError
		     AND hFileHandle <> 0
		THEN
			bDone := FALSE;
			bError := TRUE;

			enStep := eFileClose;					(* Next step *)

		ELSE
			bBusy := FALSE;
			bDone := FALSE;
			bError := TRUE;
	
			enStep := eNotExecute;					(* Next step *)
		END_IF

	eNotExecute:
		IF NOT bExecute
		THEN
			bBusy := FALSE;
			bDone := FALSE;
			bError := FALSE;
			udnErrNo := 0;

			enStep := eWaitExecute;			(* Next step *)

		END_IF

END_CASE

fbCreateDir(
	sNetId:= '',
	sPathName:= sFilePath,
	ePath:= PATH_GENERIC,
	tTimeout:= tTimeout);
fbFileOpen(
	sNetId := '',
	sPathName := sPathName,
	nMode := dwModeCache,
	ePath := PATH_GENERIC,
	tTimeout := tTimeout);
fbFileClose(
	sNetId := '',
	hFile := hFileHandle,
	tTimeout := tTimeout );
fbFileWrite(
	sNetId := '',
	hFile := hFileHandle,
	pWriteBuff := ADR(sWriteRecordCache),
	cbWriteLen := INT_TO_UDINT(LEN(sWriteRecordCache)),
	tTimeout := tTimeout);
fbFileRead(
	sNetId := '',
	hFile := hFileHandle,
	pReadBuff := ADR(sReadRecord),
	cbReadLen := INT_TO_UDINT(LEN(sReadRecord)),
	tTimeout := tTimeout);

END_FUNCTION_BLOCK

// ---- POUs/Tc3 Objects/File/TXT/FB_LoadFromFile_1.TcPOU
FUNCTION_BLOCK FB_LoadFromFile_1
(*
Function to make easier work with file. Below options to choose. 
Chose option doasn't work with the others option. Allways is checking  only exist of file.
 
00000000 - 0 - Only check exist of file.
00000001 - 1 - Read line by line and save to array of string.
00000010 - 2 - Read line by line. Save first signs to string and convert to array of bool.
00000011 - 3 - Transfer  array form file to array of string on PLC - requirements:
			- kind of columns separator (bySep) and sign end of line (byEndLine),
			- amount of rows (usiMaxDimR) and columns (usiMaxDimR) to read.
00000111 - 4 - Option 3 + filter float numer readable

Constructor: 		Patryk Panylo
Company:		E. Riexinger GmbH
Date:			18.11.2015
Version:			1.00

Date:			Revision:		Who:				Comment
dd.mm.yyyy		x.xx			Initials			comment

*)
VAR_INPUT
	(* Enummerations *)

	(* Variables *)
	bEnable						:BOOL;									(* Enable FB *)
	bExecute					:BOOL; 									(* Execute load data *)
	byConfig 					:BYTE := 0;								(* Configuration byte
																		    Options:  - 2#00000000 (default),
																				    - 2#00000001 (actOption1),
																			  	    - 2#00000010 (actOption2),
																				    - 2#00000011 (actOption3),
																				    - 2#00000111 (actOption4),
																		*)
	sFilePath					:STRING;								(* File path *)
	sFileName					:STRING;								(* File name *)
	sFileSuffix					:STRING := 'dat';							(* Suffix of file *)
	sSep						:STRING := '$T'; 							(* Seperator sign for colums *)
	sEndLine					:STRING := '$N'; 							(* End line sign for lines *)
	sComment					:STRING := '!'; 							(* End line sign for lines *)
	tTimeout					:TIME := T#1S;							(* TimeOut *)

	(* References *)

	(* Interfaces *)


	(* Instances *)

END_VAR
VAR_OUTPUT
	(* Enummerations *)

	(* Variables *)
	arsData						:ARRAY [0..GVL_FB_LoadFromFile.usnFileArrayMaxDimR] OF STRING [255];					(* Used with Option1 -  Array with read data from file in String[160] *)
	arbDataBool					:ARRAY [0..GVL_FB_LoadFromFile.usnFileArrayMaxDimR] OF BOOL;							(* Used with Option2 - Array with read data from file in Bool *)
	arsDataDimRC				:ARRAY [0..GVL_FB_LoadFromFile.usnFileArrayMaxDimR, 0..GVL_FB_LoadFromFile.usnFileArrayMaxDimC ] OF STRING [20]; 		(* Used with Option3 - Matrix with read data from file in String[160] *)
	arrDataDimRC				:ARRAY [0..GVL_FB_LoadFromFile.usnFileArrayMaxDimR, 0..GVL_FB_LoadFromFile.usnFileArrayMaxDimC ] OF REAL; 			(* Matrix with read data from file in real *)
	bDone						:BOOL;													(* Program done *)
	bBusy						:BOOL;													(* Program busy *)
	bError						:BOOL;													(* Error *)
	udnErrorNo					:UDINT;													(* Error number *)
	sErrorMsg					:STRING; 												(* Error message *)

	(* References *)

	(* Interfaces *)

	(* Instances *)

END_VAR
VAR
	(* Enummerations *)
	etLoadFromFile				:ET_LoadFromFile;								(* Load from file enum variable *)

	(* Variables *)
	dwMode						:DWORD;										(* Contains the mode in which the file is to be opened *)
	sPathName					:STRING;										(* Contains the path and filename for the file to be opened *)
	hFileHandle					:UINT;											(* File handle *)
	usnRowsCounter				:USINT; 											(* Counter of rows (lines) in a  file*)

	sDataSign					:STRING[1];										(* Read first sign from line *)
	sDataString					:STRING[GVL_FB_LoadFromFile.usnFileArrayMaxDimR];							(* Created string of sign *)
	arbyData					:ARRAY [0..GVL_FB_LoadFromFile.usnFileArrayMaxDimR] OF BYTE;					(* String into array of byte *)
	ptString 					:POINTER TO ARRAY[0..GVL_FB_LoadFromFile.usnFileArrayMaxDimR] OF BYTE;		(* Pointer to sDataString *)

	byDataSign					:BYTE;											(* Marker for sign form line *)
	ptByte						:POINTER TO BYTE;								(* Pointer to arsData *)
	usnColumnsCounter 			:USINT; 											(* Counter of colums *)

	bFirstTime					:BOOL;

	(* References *)

	(* Interfaces *)

	(* Instances *)
	tonTimeout					:TON;

	fbFileOpen					:FB_FileOpen;		(* Open file *)
	fbFileGets					:FB_FileGets;			(* Read from file *)
	fbFileClose					:FB_FileClose;		(* Close file *)

	rtExecute					:R_TRIG;				(* Positive edge for start *)

END_VAR

IF NOT bEnable
THEN
	bDone := FALSE;					(* Program done *)
	bBusy := FALSE;                                  	(* Program not busy *)
	bError := FALSE;                                 	(* Program not error *)
	udnErrorNo := 0;                                 		(* Error number *)

	bFirstTime := FALSE;
	RETURN;
END_IF;

IF NOT bFirstTime
THEN
	bDone := FALSE;                                 	(* Program done *)
	bBusy := FALSE;                                  	(* Program not busy *)
	bError := FALSE;                                 	(* Program not error *)
	udnErrorNo := 0;                                		(* Error number *)

	etLoadFromFile := ET_LoadFromFile_eWaitExecute;       				(* Next step *)
	
	bFirstTime := TRUE;
END_IF;

sPathName := CONCAT(
				sFilePath, CONCAT(
							sFileName, CONCAT(
										'.', sFileSuffix)));

rtExecute(CLK:= bExecute);				(* Positive edge for start *)

CASE etLoadFromFile OF
        
	ET_LoadFromFile_eWaitExecute:
		bBusy := FALSE;                                     		(* Program not busy *)
		bError := FALSE;                                    		(* Program not error *)

		IF rtExecute.Q
		THEN
			bDone := FALSE;                                 	(* Program done, in position *)
			bBusy := TRUE;                                  	(* Program busy *)
			udnErrorNo := 0;
			usnRowsCounter := 0;

			fbFileOpen.bExecute := FALSE;			(* File open *)
			fbFileClose.bExecute := FALSE;			(* File close *)
			fbFileGets.bExecute := FALSE;			(* File read *)

			dwMode := FOPEN_MODEREAD OR FOPEN_MODETEXT;

			etLoadFromFile := ET_LoadFromFile_eFileName;         		(* Next step *)
		END_IF;

	ET_LoadFromFile_eFileName:
		IF sFilePath <> ''
		     AND sFileName <> ''
		     AND sFileSuffix <> ''
		     AND byConfig <> 0
		THEN
			etLoadFromFile := ET_LoadFromFile_eChkFileExist;            			(* Next step *)

		ELSE
			udnErrorNo := INT_TO_UINT(ET_LoadFromFile_eFileName);

			etLoadFromFile := ET_LoadFromFile_eError;            			(* Next step *)

		END_IF

	ET_LoadFromFile_eChkFileExist:
		etLoadFromFile := ET_LoadFromFile_eFileOpen;            			(* Next step *)

	ET_LoadFromFile_eFileOpen:
		fbFileOpen.bExecute := TRUE;

		etLoadFromFile := ET_LoadFromFile_eChkFileOpen;            			(* Next step *)

	ET_LoadFromFile_eChkFileOpen:
		IF NOT fbFileOpen.bBusy
		     AND NOT fbFileOpen.bError
		THEN
			fbFileOpen.bExecute := FALSE;
			hFileHandle := fbFileOpen.hFile;

			MEMSET(ADR(arsData), 0, SIZEOF(arsData));						(* Array reset *)
			MEMSET(ADR(arbDataBool), 0, SIZEOF(arbDataBool));				(* Array reset *)
			MEMSET(ADR(arsDataDimRC), 0, SIZEOF(arsDataDimRC)); 		(* Array reset *)
			MEMSET(ADR(arrDataDimRC), 0, SIZEOF(arrDataDimRC)); 			(* Array reset *)

			etLoadFromFile := ET_LoadFromFile_eReadData;            			(* Next step *)

		ELSIF fbFileOpen.bError
		THEN
			fbFileOpen.bExecute := FALSE;
			udnErrorNo := fbFileOpen.nErrId;

			etLoadFromFile := ET_LoadFromFile_eError;            			(* Next step *)

		END_IF

	ET_LoadFromFile_eReadData:
		fbFileGets.bExecute := TRUE;

		etLoadFromFile := ET_LoadFromFile_eChkReadData;            			(* Next step *)

	ET_LoadFromFile_eChkReadData:
		IF NOT fbFileGets.bBusy
		     AND NOT fbFileGets.bError
		THEN
			fbFileGets.bExecute := FALSE;

			CASE byConfig OF
				1:	A_Option1();				(* Call option 1 *)
				2:	A_Option2();				(* Call option 2 *)
				3..4:	A_Option3();				(* Call option 3,4 *)
			END_CASE

		ELSIF fbFileGets.bError
		THEN
			fbFileGets.bExecute := FALSE;
			udnErrorNo := fbFileGets.nErrId;

			etLoadFromFile := ET_LoadFromFile_eError;            			(* Next step *)

		END_IF

	ET_LoadFromFile_eFileClose:
		fbFileClose.bExecute := TRUE;

		etLoadFromFile := ET_LoadFromFile_eChkFileClose;            			(* Next step *)

	ET_LoadFromFile_eChkFileClose:
		IF NOT fbFileClose.bBusy
		     AND NOT fbFileClose.bError
		THEN
			fbFileClose.bExecute := FALSE;

			IF NOT bError
			THEN
				etLoadFromFile := ET_LoadFromFile_eDone;            			(* Next step *)
			ELSE
				etLoadFromFile := ET_LoadFromFile_eError;            			(* Next step *)
			END_IF


		ELSIF fbFileClose.bError
		THEN
			fbFileClose.bExecute := FALSE;
			udnErrorNo := fbFileClose.nErrId;

			etLoadFromFile := ET_LoadFromFile_eError;            			(* Next step *)

		END_IF

	ET_LoadFromFile_eDone:
		bDone := TRUE;                                      		(* Program done, in position *)
		bBusy := FALSE;                                     		(* Program not busy *)
		bError := FALSE;
		udnErrorNo := 0;
	
		etLoadFromFile := ET_LoadFromFile_eNoExecute;            		(* Next step *)

	ET_LoadFromFile_eError:
		IF NOT bError
		     AND hFileHandle <> 0
		THEN
			bDone := FALSE;                                    	 	(* Program done, in position *)
			bError := TRUE;                                     		(* Program error *)
			bBusy := FALSE;                                     		(* Program not busy *)
	
			etLoadFromFile := ET_LoadFromFile_eFileClose;            		(* Next step *)

		ELSE
			bDone := FALSE;                                    	 	(* Program done, in position *)
			bError := TRUE;                                     		(* Program error *)
			bBusy := FALSE;                                     		(* Program not busy *)

			etLoadFromFile := ET_LoadFromFile_eNoExecute;            		(* Next step *)
		END_IF

	ET_LoadFromFile_eNoExecute:
		IF NOT bExecute
		THEN
			bDone := FALSE;                                 	(* Program done *)
			bBusy := FALSE;                                 	(* Program not busy *)
			bError := FALSE;                                		(* Program not error *)
			udnErrorNo := 0;
	
			etLoadFromFile := ET_LoadFromFile_eWaitExecute;       		(* Next step *)
	
		END_IF;
        
END_CASE;

fbFileOpen(
	sNetId := '',
	sPathName := sPathName,
	nMode := dwMode,
	ePath := PATH_GENERIC,
	tTimeout := tTimeout
);
fbFileClose(
	sNetId := '',
	hFile := hFileHandle,
	tTimeout := tTimeout
);

fbFileGets(
	sNetId := '',
	hFile :=  hFileHandle,
	tTimeout := tTimeout
);

ACTION A_Option1:
(* Option 1:

00000001 - 1 - Read line by line and save to array of string.

*)
(*****************************************************************************************************************************************************************************************************)

arsData[usnRowsCounter] := fbFileGets.sLine;											(* Read line (255 chars) from file *)

IF NOT fbFileGets.bEOF															(* Check received all data form file *)
THEN
	usnRowsCounter := usnRowsCounter + 1;
	etLoadFromFile := ET_LoadFromFile_eReadData;  									(* Read next line form file *)

ELSE
	etLoadFromFile := ET_LoadFromFile_eFileClose;  									(* Close current file *)

END_IF
END_ACTION

ACTION A_Option2:
(* Option 2:

00000010 - 2 - Read line by line. Save first signs to string and convert to array of bool.

*)
(*****************************************************************************************************************************************************************************************************)

sDataSign := fbFileGets.sLine;														(* Read first sign from line *)
sDataString := CONCAT(sDataString, sDataSign);										(* Created string of sign *)

ptString := ADR(sDataString);														(* Take adress to pointer of byte *)
arbyData :=  ptString^;																(* Take string into array of byte *)
arbDataBool[usnRowsCounter] := BYTE_TO_BOOL(arbyData[usnRowsCounter] AND 16#01);	(* Move data to Array of Bool *)

IF NOT fbFileGets.bEOF															(* Check received all data form file *)
THEN
	usnRowsCounter := usnRowsCounter + 1;
	etLoadFromFile := ET_LoadFromFile_eReadData;  									(* Read next line form file *)

ELSE
	etLoadFromFile := ET_LoadFromFile_eFileClose;  									(* Close current file *)

END_IF
END_ACTION

ACTION A_Option3:
(*Option 3:

00000011 - 3 - Transfer  array form file to array of string on PLC - requirements:
			- kind of columns separator (bySep) and sign end of line (byEndLine),
			- amount of rows (usiMaxDimR) and columns (usiMaxDimR) to read.

*)
(*****************************************************************************************************************************************************************************************************)

IF usnRowsCounter <= usnFileArrayMaxDimR 							(* Choose amount of rows from file *)
    AND NOT fbFileGets.bEOF
THEN
	arsData[usnRowsCounter] := fbFileGets.sLine; 						(* Read line (255 chars) from file *)

	ptByte := ADR(arsData[usnRowsCounter]);
	byDataSign :=  ptByte^;

	usnColumnsCounter := 0;
	REPEAT

		WHILE byDataSign <> F_ToASC(sSep) 			(* $T = HEX 09 *)   (* ; = HEX 3B *) (* EOF *)	(* Reaction for special sign in string*)
			  AND  byDataSign <> F_ToASC(sEndLine)	(* $N = HEX 0A *)
		DO
			IF byDataSign = F_ToASC(sComment)
			   //OR byDataSign = F_ToASC('i')
			THEN
				EXIT;
			END_IF

			arsDataDimRC[usnRowsCounter , usnColumnsCounter] := CONCAT(arsDataDimRC[usnRowsCounter , usnColumnsCounter], F_ToCHR(byDataSign)); 	(* Read sign and create string*)

			ptByte := ptByte + 1;
			byDataSign :=  ptByte^;

		END_WHILE

		IF byConfig = 4
		THEN
			IF F_CheckStringIsReal(arsDataDimRC[usnRowsCounter , usnColumnsCounter])
			THEN
				arrDataDimRC[usnRowsCounter , usnColumnsCounter] :=  STRING_TO_REAL(arsDataDimRC[usnRowsCounter , usnColumnsCounter]);				(* Create real *)
			ELSE
				udnErrorNo := 31;

				etLoadFromFile := ET_LoadFromFile_eError;            			(* Next step *)
				RETURN;
			END_IF
		END_IF
		
		IF byDataSign <> F_ToASC(sEndLine)					(* Check end of line *)
		THEN
			IF byDataSign = F_ToASC(sComment)
			THEN
				EXIT;
			END_IF

			usnColumnsCounter := usnColumnsCounter + 1;			(* Set next columns *)
			ptByte := ptByte + 1;
			byDataSign :=  ptByte^;

		END_IF

	UNTIL byDataSign  = F_ToASC(sEndLine)					(* End when founds the end line sign*)
	END_REPEAT

	IF byDataSign <> F_ToASC(sComment)
	THEN
		usnRowsCounter := usnRowsCounter + 1;
	END_IF

	etLoadFromFile := ET_LoadFromFile_eReadData;  									(* Read next line form file *)

ELSE
	etLoadFromFile := ET_LoadFromFile_eFileClose;  									(* Close current file *)

END_IF
END_ACTION

END_FUNCTION_BLOCK

// ---- POUs/Tc3 Objects/Logger/FB_LoggerFile_1.TcPOU
FUNCTION_BLOCK FB_LoggerFile_1
(*

This function block is used to write loggin datas into file.

Constructor: 		Patryk Panylo
Company:		E. Riexinger GmbH
Date:			25.03.2014
Version:			1.00

Date:			Revision:		Who:				Comment
dd.mm.yyyy		x.xx			Initials			comment

*)

VAR_INPUT
	bEnable						:BOOL;					(* Enable FB *)
	bExecute					:BOOL;					(* Execute operation *)
	sFilePath					:STRING;				(* File path *)
	sFileName					:STRING;				(* File name *)
	sFileSuffix					:STRING := 'dat';			(* Suffix of file *)
	arstLoggerWaitInterrupt			:ARRAY[1..GVL_Logger.unLOG_BEFOR_MAX_NO] OF ST_LoggerVar;			(* Data to write to file *)
	arstLoggerDuringInterrupt		:ARRAY[1..GVL_Logger.unLOG_DURING_MAX_NO] OF ST_LoggerVar;			(* Data to write to file *)
	arstLoggerAfterInterrupt			:ARRAY[1..GVL_Logger.unLOG_AFTER_MAX_NO] OF ST_LoggerVar;			(* Data to write to file *)
	tTimeout						:TIME := t#1s;				(* States the time before the function is cancelled *)
END_VAR
VAR_OUTPUT
	bBusy						:BOOL;					(* Program busy *)
	bDone						:BOOL;					(* Program done *)
	bError						:BOOL;					(* Program error *)
	udnErrNo					:UDINT;					(* Error number *)
END_VAR
VAR_IN_OUT

END_VAR
VAR
	(* Enummerations *)
	enStep						: (eWaitExecute := 0, eChkFileName, eChkeNumOfRecords, eFileOpen, eChkFileOpen, eFilePuts, eChkFilePuts, eFileClose, eChkFileClose, eDone, eError, eNotExecute);			(* Sequence state for open, read/write and close the file *)
	enGetData					: (eWaitInterruptData, eDuringInterruptData, eAfterInterruptData, eNoData);					(* Sequence state for data *)

	(* Variables *)
	bFirstTime					:BOOL;					(* First PLC cycle *)
	unLogSize					:UINT;
	unLogIdx						:UINT;
	unRecordsSize				:UINT;
	unRecordsIdx					:UINT;

	dwMode						:DWORD;				(* Contains the mode in which the file is to be opened *)
	sPathName					:STRING;				(* Contains the path and filename for the file to be opened *)
	hFileHandle					:UINT;					(* File handle *)

	unPutsCounter				:UINT;

	sRecordsToWrite				:STRING;

	(* Instances *)
	fbFileOpen					:FB_FileOpen;			(* File open *)
	fbFileClose					:FB_FileClose;			(* File close *)
	fbFilePuts					:FB_FilePuts;				(* File puts *)

END_VAR
VAR CONSTANT
	sSeparator					:STRING := '$T';
	sNewLine					:STRING := '$N'; 							(* End line sign for lines *)
END_VAR

IF NOT bEnable				(* Enable FB *)
THEN
	bFirstTime := FALSE;		(* First PLC cycle *)
	bBusy := FALSE;			(* Program busy *)
	bDone := FALSE;			(* Program done *)
	bError := FALSE;			(* Program error *)
	udnErrNo := 0;				(* Error number *)
	RETURN;
END_IF

IF NOT bFirstTime
THEN
	bBusy := FALSE;			(* Program busy *)
	bDone := FALSE;			(* Program done *)
	bError := FALSE;			(* Program error *)

	enStep := eWaitExecute;

	bFirstTime := TRUE;
END_IF


(* Sequence state for open, read/write and close the file *)
CASE enStep
OF

	eWaitExecute:
		IF bExecute
		THEN
			fbFileOpen.bExecute := FALSE;			(* File open *)
			fbFileClose.bExecute := FALSE;			(* File close *)
			fbFilePuts.bExecute := FALSE;			(* File puts *)

			bBusy := TRUE;
			bDone := FALSE;
			bError := FALSE;
			udnErrNo := 0;

			dwMode := FOPEN_MODEWRITE OR FOPEN_MODETEXT;

			enStep := eChkFileName;			(* Next step *)

		END_IF

	(* Check file name and path *)
	eChkFileName:

		sPathName := CONCAT(
						sFilePath, CONCAT(
									sFileName, CONCAT(
												'.', sFileSuffix)));

		IF sFilePath <> ''
		     AND sFileName <> ''
		     AND sFileSuffix <> ''
		THEN
			enStep := eChkeNumOfRecords;			(* Next step *)

		ELSE
			udnErrNo := eChkFileName;

			enStep := eError;				(* Next step *)

		END_IF

	(* Check number of records to save *)
	eChkeNumOfRecords:
		IF GVL_Logger.unNUM_OF_LOG_VAR = 0
		THEN
			enStep := eDone;				(* Next step *)
	
		ELSE
			enStep := eFileOpen;			(* Next step *)

		END_IF
	(* Open the file *)
	eFileOpen:
		fbFileOpen.bExecute := TRUE;

		enStep := eChkFileOpen;				(* Next step *)

	(* Check open the file *)
	eChkFileOpen:
		IF NOT fbFileOpen.bBusy
		THEN
			IF NOT fbFileOpen.bError
			THEN
				fbFileOpen.bExecute := FALSE;
				hFileHandle := fbFileOpen.hFile;

				unLogIdx := 0;
		  		unRecordsIdx := 0;

				enGetData := eWaitInterruptData;
				enStep := eFilePuts;			(* Next step *)

			ELSE
				fbFileOpen.bExecute := FALSE;
				udnErrNo := fbFileOpen.nErrId;
	
				enStep := eError;					(* Next step *)

			END_IF
		END_IF

	(* Puts data into the file *)
	eFilePuts:
		(* Get data *)
		A_GetData();

		IF LEN(sRecordsToWrite) > 254
		THEN
			sRecordsToWrite := DELETE(
								sRecordsToWrite,
								LEN(sRecordsToWrite) + 1 - 254, 254
							    );
		END_IF


		sRecordsToWrite := CONCAT(
							sRecordsToWrite,
							SEL(unRecordsIdx = 0, sSeparator, sNewLine)
						    );


		fbFilePuts.bExecute := TRUE;

		enStep := eChkFilePuts;				(* Next step *)

	(* Check puts the file *)
	eChkFilePuts:
		IF NOT fbFilePuts.bBusy
		THEN
			IF NOT fbFilePuts.bError
			THEN
				fbFilePuts.bExecute := FALSE;
				unPutsCounter := unPutsCounter + 1;

				IF enGetData = eNoData
				THEN
					enStep := eFileClose;				(* Next step *)
				ELSE
					enStep := eFilePuts;				(* Next step *)
				END_IF

			ELSIF  fbFilePuts.bError
			THEN
				fbFilePuts.bExecute := FALSE;
				udnErrNo := fbFilePuts.nErrId;

				enStep := eError;					(* Next step *)

			END_IF
		END_IF

	(* Close the file *)
	eFileClose:
		fbFileClose.bExecute := TRUE;

		enStep := eChkFileClose;				(* Next step *)

	(* Check close the file *)
	eChkFileClose:
		IF NOT fbFileClose.bBusy
		THEN
			IF NOT fbFileClose.bError
			THEN
				fbFileClose.bExecute := FALSE;
				enStep := eDone;					(* Next step *)

				IF bError
				THEN
					enStep := eError;				(* Next step *)
				END_IF

			ELSE
				fbFileClose.bExecute := FALSE;
				udnErrNo := fbFileClose.nErrId;
	
				enStep := eError;					(* Next step *)
				
			END_IF
		END_IF

	eDone:
		bBusy := FALSE;
		bDone := TRUE;
		bError := FALSE;
		udnErrNo := 0;

		enStep := eNotExecute;					(* Next step *)

	eError:
		IF NOT bError
		     AND hFileHandle <> 0
		THEN
			bDone := FALSE;
			bError := TRUE;

			enStep := eFileClose;					(* Next step *)

		ELSE
			bBusy := FALSE;
			bDone := FALSE;
			bError := TRUE;
	
			enStep := eNotExecute;					(* Next step *)
		END_IF

	eNotExecute:
		IF NOT bExecute
		THEN
			bBusy := FALSE;
			bDone := FALSE;
			bError := FALSE;
			udnErrNo := 0;

			enStep := eWaitExecute;			(* Next step *)

		END_IF

END_CASE

fbFileOpen(
	sNetId := '',
	sPathName := sPathName,
	nMode := dwMode,
	ePath := PATH_GENERIC,
	tTimeout := tTimeout
);
fbFileClose(
	sNetId := '',
	hFile := hFileHandle,
	tTimeout := tTimeout
);
fbFilePuts(
	sNetId := '',
	hFile:= hFileHandle,
	sLine := sRecordsToWrite,
	tTimeout := tTimeout
 );

ACTION A_GetData:

CASE enGetData
OF
	eWaitInterruptData:
		IF unLogIdx = 0
		THEN
			unLogIdx := 1;
			unLogSize := unLOG_BEFOR_MAX_NO;

			sRecordsToWrite := '[WAIT INTERRUPT]';

		ELSIF unRecordsIdx = 0
		THEN
			unRecordsIdx	 := 1;
			unRecordsSize := unNUM_OF_LOG_VAR;

			sRecordsToWrite := CONCAT(
								UDINT_TO_STRING(arstLoggerWaitInterrupt[unLogIdx].udnCycleNo),
								CONCAT(
									sSeparator,
									arstLoggerWaitInterrupt[unLogIdx].sTimeStamp
								)
							   );

		ELSE

			sRecordsToWrite := arstLoggerWaitInterrupt[unLogIdx].arsLogVars[unRecordsIdx];

			unRecordsIdx := unRecordsIdx + 1;

			IF unRecordsIdx > unRecordsSize
			THEN
				unRecordsIdx := 0;
				unLogIdx := unLogIdx + 1;
			END_IF

		END_IF

		IF unLogIdx > unLogSize
		THEN
			unLogIdx := 0;
		  	unRecordsIdx := 0;
			enGetData := eDuringInterruptData;					(* Next step *)
		END_IF

	eDuringInterruptData:

		IF unLogIdx = 0
		THEN
			unLogIdx := 1;
			unLogSize := unLOG_DURING_MAX_NO;

			sRecordsToWrite := '[DURING INTERRUPT]';

		ELSIF unRecordsIdx = 0
		THEN
			unRecordsIdx	 := 1;
			unRecordsSize := unNUM_OF_LOG_VAR;

			sRecordsToWrite := CONCAT(
								UDINT_TO_STRING(arstLoggerDuringInterrupt[unLogIdx].udnCycleNo),
								CONCAT(
									sSeparator,
									arstLoggerDuringInterrupt[unLogIdx].sTimeStamp
								)
							   );

		ELSE
			sRecordsToWrite := arstLoggerDuringInterrupt[unLogIdx].arsLogVars[unRecordsIdx];

			unRecordsIdx := unRecordsIdx + 1;

			IF unRecordsIdx > unRecordsSize
			THEN
				unRecordsIdx := 0;
				unLogIdx := unLogIdx + 1;
			END_IF

		END_IF

		IF unLogIdx > unLogSize
		THEN
			unLogIdx := 0;
		  	unRecordsIdx := 0;
			enGetData := eAfterInterruptData;					(* Next step *)
		END_IF

	eAfterInterruptData:

		IF unLogIdx = 0
		THEN
			unLogIdx := 1;
			unLogSize := unLOG_AFTER_MAX_NO;

			sRecordsToWrite := '[AFTER INTERRUPT]';

			IF LEN(arstLoggerAfterInterrupt[unLogIdx].sTimeStamp) = 0
			THEN
				unLogIdx := GVL_Logger.unLOG_AFTER_MAX_NO + 1;
			END_IF

		ELSIF unRecordsIdx = 0
		THEN
			unRecordsIdx	 := 1;
			unRecordsSize := unNUM_OF_LOG_VAR;

			sRecordsToWrite := CONCAT(
								UDINT_TO_STRING(arstLoggerAfterInterrupt[unLogIdx].udnCycleNo),
								CONCAT(
									sSeparator,
									arstLoggerAfterInterrupt[unLogIdx].sTimeStamp
								)
							   );

		ELSE
			sRecordsToWrite := arstLoggerAfterInterrupt[unLogIdx].arsLogVars[unRecordsIdx];

			unRecordsIdx := unRecordsIdx + 1;

			IF unRecordsIdx > unRecordsSize
			THEN
				unRecordsIdx := 0;
				unLogIdx := unLogIdx + 1;
			END_IF

		END_IF

		IF unLogIdx > unLogSize
		THEN
			unLogIdx := 0;
		  	unRecordsIdx := 0;
			enGetData := eNoData;
		END_IF

	eNoData:
		unLogIdx := 0;
		 unRecordsIdx := 0;

END_CASE
END_ACTION

END_FUNCTION_BLOCK

// ---- POUs/Tc3 Objects/Logger/FB_Logger_1.TcPOU
FUNCTION_BLOCK FB_Logger_1
VAR_INPUT
	bEnable								:BOOL;
	bEnableSaveInFile					:BOOL;				(* Enable save in file *)
	bInterrupt							:BOOL;
	sDateTime 							:STRING;			(* Actual date and time *)
	bDeleteAll							:BOOL;
	bLogOne								:BOOL := FALSE;		(* Log data only one time *)
	sFilePath							:STRING := 'C:\TwinCAT\Boot\';			(* Login file path *)
	sFileSuffix							:STRING := 'log';							(* Suffix of loggin file *)
	arsLogVars							:ARRAY[1..GVL_Logger.unNUM_OF_LOG_VAR] OF STRING(10);
	unLogMaxNo							:UINT;
	unLogBeforMaxNo						:UINT;
	unLogDuringMaxNo					:UINT;
	unLogAfterMaxNo						:UINT;
END_VAR
VAR_OUTPUT
	bBusy								:BOOL;
	bDone								:BOOL;
	bError								:BOOL;
	bEStop								:BOOL;
	arstLogger							:ARRAY[1..GVL_Logger.unLOG_MAX_NO] OF ST_Logger;
	arstLoggerWaitInterrupt				:ARRAY[1..GVL_Logger.unLOG_BEFOR_MAX_NO] OF ST_LoggerVar;
	arstLoggerDuringInterrupt			:ARRAY[1..GVL_Logger.unLOG_DURING_MAX_NO] OF ST_LoggerVar;
	arstLoggerAfterInterrupt			:ARRAY[1..GVL_Logger.unLOG_AFTER_MAX_NO] OF ST_LoggerVar;
END_VAR
VAR
	bFirstTime							:BOOL;
	nIdx								:INT;			(* Index *)
	udnCycleNo							:UDINT;
	unInstanceIdx						:UINT;

	unState								:UINT := 0;
	unIncLog							:UINT := 1;
	unIncDuringInterrupt				:UINT := 1;
	unIncAfterInterrupt					:UINT := 1;

	rtDeleteAll							:R_TRIG;
	rtInterrupt							:R_TRIG;
	fbLoggerFile						:FB_LoggerFile;

